(* IEC 61131-3 sources: 89152_FlorisHendrix_AfstudeerProject/89152_FlorisHendrix_ExamenProject/Stations/MachineControl/MachineControl/Class/HwControl, 1 file *)

(* ---- HwControl.st ---- *)
#include "..\..\Class\HwControl\HwControl.h"
#include "..\..\Class\HwControl\watchdog.h"
#include "..\..\Source\interfaces\lsl_st_sysinfo.h"
#include "..\..\Source\interfaces\lsl_st_systrace.h"
#include "..\..\Class\HwControl\_HWKScope.h"

(*!
<Class
	Name               = "HwControl"
	Revision           = "5.21"
	RealtimeTask       = "false"
	DefRealtime        = "1 ms"
	DefRealtimeIndex   = "0"
	CyclicTask         = "false"
	DefCyclictime      = "1 ms"
	DefCyclicIndex     = "2147483392"
	BackgroundTask     = "false"
	Sigmatek           = "true"
	OSInterface        = "false"
	HighPriority       = "false"
	Automatic          = "false"
	UpdateMode         = "Prescan"
	IconPath           = ".\Class\HwControl\HwControl.ico"
	SharedCommandTable = "true"
	Objectsize         = "(646,120)"
	Comment            = "Class to handle VaranManager,  and the cooperation with DiasMasterC">
	<Channels>
		<Server Name="Control">
		</Server>
		<Server Name="DiasMaster" WriteProtected="false" Comment="connect to client &apos;to_HWControl&quot; of class DiasMasterC if used (if Server is 1 class is connected)&#13;&#10;">
		</Server>
		<Server Name="SafetyState" Visualized="true" Initialize="false" WriteProtected="true" Retentive="false" Comment="Shows state of safety functionality initialisation&#13;&#10;&#13;&#10; 1..OK&#13;&#10; 0..not active or initializing&#13;&#10;-1..failed to allocate memory&#13;&#10;-2..invalid domain number set in this system&#13;&#10;-3..newer OS version required for domain number support&#13;&#10;-4..method to determine domain number not provided by lsl_st_hardwaretree.h&#13;&#10;-5..only 1 instance of safety manager allowed&#13;&#10;-6..a slave system can only have 1 master. check hw class configuration&#13;&#10;-7..invalid module type tried to log in&#13;&#10;-8..couldn&apos;t find InterfaceCRC which is requested by other domain. Check SafetyDesigner projects, most likely the interface variables doesn&apos;t match.&#13;&#10;-9..failed to add a new copy data object to varan manager&#13;&#10;-10..a non-optional module or domain is not available&#13;&#10;-11..timeout in initialisation (see debugger trace or logfile for further details)&#13;&#10;-13..the class safetymanager could not login into the class HwControl."/>
		<Client Name="HwcLogging" Required="true" Internal="true"/>
		<Client Name="HWRtPostScan" Required="true" Internal="true"/>
		<Client Name="InterfaceNo" Required="false" Internal="false" DefValue="1" Comment="If interface frames via IP address are used, this is the place to choose the interface number&#13;&#10;&#13;&#10;For example if you set the IP of interface 1 via autoexec.lsl setting SET IP 1 HOSTADDR x.x.x.x and this is what you want to use, you choose 1 for the interface number."/>
		<Client Name="RtTaskSync" Required="false" Internal="false" DefValue="0" Comment="With this setting the realtime task synchronization between more cores can be activated.&#13;&#10;If it is activated and not supported, the client is set to 0.&#13;&#10;As an initialization value. For further information look at library help.&#13;&#10;0 .. deactivated (default)&#13;&#10;1 .. activated&#13;&#10;&#13;&#10;"/>
		<Client Name="SafetyDomainTimeout" Required="false" Internal="false" Comment="[ms] the class has to wait for optional interface domains (leave 0 if none available)&#13;&#10;Set this client to 1 when using FlexCon functionality (without interface domains) where it&apos;s possible that not all participants are available at all times"/>
		<Client Name="SafetyManager" Required="true" Internal="true"/>
		<Client Name="UdpSafetyPort" Required="false" Internal="false" DefValue="10823" Comment="If interface frames via IP address are used, this is the place to choose the port.&#13;&#10;It&apos;s recommended to only change the port (all communication partners must use the same port!) if there would be a conflict with the default port 10823."/>
	</Channels>
	<Dependencies>
		<Files>
			<File Path=".\Class\VaranManager_Base\VaranManager_Base.h" Include="false"/>
			<File Path=".\Class\HwControl\HwControl.h" Include="true"/>
			<File Path=".\Class\HwControl\watchdog.h" Include="true"/>
			<File Path=".\Source\interfaces\lsl_st_sysinfo.h" Include="true"/>
			<File Path=".\Source\interfaces\lsl_st_systrace.h" Include="true"/>
			<File Path=".\Class\HwControl\_HWKScope.h" Include="true"/>
		</Files>
	</Dependencies>
	<RevDoku>
		<Owner Company="Sigmatek" Author="renste"/>
		<Dokumentation Revision="5.21" Date="30.09.2022" Author="RamAnd" Company="Sigmatek" Description="The busy state of the safety CPU wasn&apos;t detected correctly when establishing UDP connections."/>
		<Dokumentation Revision="5.20" Date="13.07.2022" Author="RamAnd" Company="Sigmatek" Description="Try again to establish a safety UDP connection if the attempt failed because the safe CPU was busy."/>
		<Dokumentation Revision="5.19" Date="22.03.2022" Author="RamAnd" Company="Sigmatek" Description="Added support for the new OS Interface to quit errors"/>
		<Dokumentation Revision="5.18" Date="17.01.2022" Author="EisMic" Company="Sigmatek" Description="Testversion: Forward the NewInst commando CMD_HWC_CONVERT_COMPRESSED_HWPATH to the SafetyManager class."/>
		<Dokumentation Revision="5.17" Date="30.11.2021" Author="EisMic" Company="Sigmatek" Description="Added global functions to determine the current operation system.&#13;&#10;Added global function HWC_IsPostInitFinished to determine if the postinit phase is finished or not."/>
		<Dokumentation Revision="5.16" Date="23.10.2020" Author="PieSte" Company="Sigmatek" Description="Added support for new blocktype and extended routing of FSoE data for this type.&#13;&#10;Corrected allocate of udp buffers at &quot;AddModule()&quot;.&#13;&#10;Don&apos;t Log AddDynSlave error if RetCode is zero at GetDestSafetyOfDO() Methode."/>
		<Dokumentation Revision="5.15" Date="18.12.2020" Author="RamAnd" Company="Sigmatek" Description="Removed CLI/STI occurances in internal time measurements"/>
		<Dokumentation Revision="5.14" Date="13.03.2020" Author="Berste1" Company="Sigmatek" Description="Registration for Pll readjustment added"/>
		<Dokumentation Revision="5.13" Date="08.04.2020" Author="PieSte" Company="Sigmatek" Description="Add client RtTaskSync for realtime synchronization if more than one core is used.&#13;&#10;Corrected nil pointer &quot;pStr_HWTreeEntry&quot; at newinst command &quot;CMD_GET_HARDWARE_DIAGNOSIS&quot;."/>
		<Dokumentation Revision="5.12" Date="02.03.2020" Author="FurDom" Company="Sigmatek" Description="Reworked to support newer CPUs (address space &gt; 0x80000000). Needs SafetyUDP class version &gt;= 1.4!"/>
		<Dokumentation Revision="5.11" Date="14.08.2019" Author="LanSte" Company="Sigmatek" Description="Added header file: _HWKScope.h for scope interface. "/>
		<Dokumentation Revision="5.10" Date="08.11.2019" Author="RamAnd" Company="Sigmatek" Description="Detached the logging functionality from HwControl into a new class HwcLogging which is used now as an embedded object in HwControl.&#13;&#10;Added more logging possibilities via new function _HwcLog_sprintfST."/>
		<Dokumentation Revision="5.9" Date="18.07.2019" Author="RamAnd" Company="Sigmatek" Description="Corrected that SDO forwarding would not work properly in some cases.&#13;&#10;Prevent writing to an invalid pointer when resetting UDP connections that could have lead to a crash."/>
		<Dokumentation Revision="5.8" Date="25.06.2019" Author="RamAnd" Company="Sigmatek" Description="Added support for FlexCon functionality."/>
		<Dokumentation Revision="5.7" Date="14.03.2019" Author="RamAnd" Company="Sigmatek" Description="Removed limitations of formerly unallowed safety topologies (since v4.0)"/>
		<Dokumentation Revision="5.6" Date="12.02.2019" Author="PieSte" Company="Sigmatek" Description="The Sequence Number in the SafetyManager class for Udp Safety communication has been extended from 1 to 4 bytes. This increases the availability of the Udp Safety connection. Furthermore two clients have been added at internal class SafetyManager to set the Request Cycle (Default 10) and the Response Timeout (Default 100ms) to optimize the Safety UDP bus load. This setting may only be changed after consultation with Sigmatek.  (SA43141)&quot;/&gt;"/>
		<Dokumentation Revision="5.5" Date="22.01.2019" Author="EisMic" Company="Sigmatek" Description="Corrected an error that the Realtime/Cyclic task of the class was called 2 times if the derivation of the class has a configured Realtime/Cyclic Task. (The error apperared since v5.0)"/>
		<Dokumentation Revision="5.4" Date="15.11.2018" Author="LanSte" Company="Sigmatek" Description="SafetyManager: Added support for custom FSoE Connections."/>
		<Dokumentation Revision="5.3" Date="27.08.2018" Author="PieSte" Company="Sigmatek" Description="Behaviour of safety udp communication when resetting the bSequenceCntReceived flag after maximum of retries corrected. (SafetyManager)"/>
		<Dokumentation Revision="5.2" Date="18.07.2018" Author="PieSte&#13;&#10;EisMic" Company="Sigmatek" Description="Added support for HGW1033-3. (in SafetyManager)&#13;&#10;Removed incorrect LogMessage. Corrected access exception in method CalculateTaskInfo.&#13;&#10;OS_AddTraceKeyVal is not used anymore with OS-Version between 9.1.0 and 9.3.0. Not supported with these versions."/>
		<Dokumentation Revision="5.1" Date="19.06.2018" Author="ZoePat" Company="Sigmatek" Description="Corrected a possible reboot of some CPUs (CCP512, CCP612, CP212, and similar). The error appeared since V5.0 if the SRAM was accessed via the cyclic-task of the HWControl."/>
		<Dokumentation Revision="5.0" Date="26.03.2018" Author="EisMic" Company="Sigmatek" Description="Added support for 2nd realtime.&#13;&#10;Added support for 2nd varanmanager.&#13;&#10;Removed task settings from object. Task-settings for realtime and cyclic task are now calculated depending on the connected hardware-classes. See documentation for more details.&#13;&#10;Extended the methods AddFirstCallHw and AddHwObject by some parameters to select a CPU-core and task-times.&#13;&#10;Added support for SmartIO modules."/>
		<Dokumentation Revision="4.15" Date="06.03.2018" Author="EisMic" Company="Sigmatek" Description="Attached header files no longer point to the installation directory of LASAL but instead now point to the the source/interfaces folder."/>
		<Dokumentation Revision="4.14" Date="18.01.2018" Author="EisMic" Company="Sigmatek" Description="Added new NewInst command to get supported features by HwControl.&#13;&#10;The newinst cmd CMD_SET_POSTINIT_DONE will now be send to all connected classes instead of only to the DiasMaster."/>
		<Dokumentation Revision="4.13" Date="23.01.2018" Author="RamAnd" Company="Sigmatek" Description="Log messages have been standardized for easier maintenance, easier use in any class and to allow spam filtering. Code for the logging functions is now only located in HwControl."/>
		<Dokumentation Revision="4.12" Date="05.01.2018" Author="PieSte" Company="Sigmatek" Description="The safety UDP communication at &quot;SafetyManager&quot; class has been made more reliable. Now only new packages are allowed and old packages are discarded."/>
		<Dokumentation Revision="4.11" Date="18.09.2017" Author="LanSte" Company="Sigmatek" Description="Added NewInst Commands to check if the Post-Init is done."/>
		<Dokumentation Revision="4.10" Date="29.08.2017" Author="RamAnd" Company="Sigmatek" Description="The VaranManager can now tell the HwControl if it doesn&apos;t have any clients connected. In this case the HwControl is in charge of triggering the internal watchdog."/>
		<Dokumentation Revision="4.9" Date="22.08.2017" Author="RamAnd" Company="Sigmatek" Description="Fixed an error which prevented two SCP111s on the same PLC from exchanging interfaceframes in both directions."/>
		<Dokumentation Revision="4.8" Date="23.05.2017" Author="RamAnd" Company="Sigmatek" Description="A pointer for dynamic parameters has been added to the hardware diagnosis. Added initialisation of the pointer with NIL."/>
		<Dokumentation Revision="4.7" Date="22.06.2017" Author="RamAnd" Company="Sigmatek" Description="If a disconnect happens in a multi master system with safety communication (more than 2 systems connected and exchanging safety data) now the other masters are notified about it to reestablish the connection."/>
		<Dokumentation Revision="4.6" Date="01.03.2017" Author="EisMic" Company="Sigmatek" Description="Corrected an error in the handling of optional safety modules."/>
		<Dokumentation Revision="4.5" Date="14.02.2017" Author="ZoePat" Company="Sigmatek" Description="SdiasModules can now request to increase the PostInit timeout."/>
		<Dokumentation Revision="4.4" Date="21.09.2016" Author="PieSte" Company="Sigmatek" Description="Add methode &quot;AddFirstCallHW&quot; for objects which are called as first at HwControl Realtime. In the TraceView scope is the and of first object call as UserEvent0 with data = 1.215.775.599 marked. "/>
		<Dokumentation Revision="4.3" Date="28.01.2016" Author="RamAnd" Company="Sigmatek" Description="Support for FSoE via IP added."/>
		<Dokumentation Revision="4.2" Date="06.06.2016" Author="EisMic" Company="Sigmatek" Description="Corrected error if distributed safety modules are connected after the initialisation phase."/>
		<Dokumentation Revision="4.1" Date="11.05.2016" Author="RamAnd" Company="Sigmatek" Description="Suppressed warning that would occur with target ARM on compiler version 30 or higher."/>
		<Dokumentation Revision="4.0" Date="30.11.2015" Author="ZoePat&#13;&#10;LanSte" Company="Sigmatek" Description="Check for unallowed safety topology."/>
		<Dokumentation Revision="3.9" Date="21.10.2015" Author="RamAnd" Company="Sigmatek" Description="Support for MS012 added"/>
		<Dokumentation Revision="3.8" Date="19.05.2015" Author="RamAnd" Company="Sigmatek" Description="If two systems with FSoE safety were connected via VBC/VMC an error in the connection establishment could cause the FSoE connection to fail."/>
		<Dokumentation Revision="3.7" Date="15.04.2015" Author="RamAnd" Company="Sigmatek" Description="Added another step in initialisation to prevent watchdog error."/>
		<Dokumentation Revision="3.6" Date="16.10.2014&#13;&#10;25.03.2015" Author="RamAnd&#13;&#10;PieSte" Company="Sigmatek" Description="Support for SCP111 added.&#13;&#10;Support for SDD1300, SDD1400, SDD1500 and SDD1600 added."/>
		<Dokumentation Revision="3.5" Date="12.11.2014" Author="PieSte" Company="Sigmatek" Description="Removed trace message if watchdog interface is not available."/>
		<Dokumentation Revision="3.4" Date="28.10.2014" Author="RamAnd" Company="Sigmatek" Description="If an error has been reported to HwControl, it is now forwarded to the DiasMasterC object (if there is one)."/>
		<Dokumentation Revision="3.3" Date="10.10.2014" Author="PieSte" Company="Sigmatek" Description="Added Watchdog API and trigger watchdog in postscan task."/>
		<Dokumentation Revision="3.2" Date="18.06.2014" Author="EisMic" Company="Sigmatek" Description="Added support for reading hardware diagnosis via newinst cmd: CMD_GET_HARDWARE_DIAGNOSE "/>
		<Dokumentation Revision="3.1" Date="17.06.2014" Author="RamAnd" Company="Sigmatek" Description="Added possibility to start a quit error via OS interface."/>
		<Dokumentation Revision="3.0" Date="15.04.2014" Author="RamAnd" Company="Sigmatek" Description="Changed initialisation: &#13;&#10; - Activation of hardware classes realtime task as well as completing CDIAS/DIAS initialisation is now done in post init instead of last init&#13;&#10; - No realtime is running in the first initialisation of the modules&#13;&#10; - New second initialisation where realtime is running to check if the realtime data are valid"/>
		<Dokumentation Revision="2.0" Date="12.02.2014" Author="PieSte" Company="Sigmatek" Description="Improved description of CyWork method."/>
		<Dokumentation Revision="1.50" Date="06.12.2013" Author="LanSte&#13;&#10;RamAnd&#13;&#10;FucHer" Company="Sigmatek" Description="Ensured that he class is copatible with old loader versions that do not support the post init phase.&#13;&#10;Removed domain support&#13;&#10;Changed AWL code to Structured Text.&#13;&#10;If the task setting for cyclic task fails, the error wasn&apos;t displayed.&#13;&#10;The task setting for cyclic task didn&apos;t work (only required if existing object is updated)."/>
		<Dokumentation Revision="1.40" Date="01.08.2013" Author="RamAnd" Company="Sigmatek" Description="Corrected error, where the user classes are already called during SDIAS initialisation."/>
		<Dokumentation Revision="1.30" Date="18.07.2013" Author="RamAnd" Company="Sigmatek" Description="Added PostInit interface of loader, where after the last init the varan managers can initialize modules until they are ready."/>
		<Dokumentation Revision="1.20" Date="07.03.2013" Author="RamAnd" Company="Sigmatek" Description="Changed range of the safety NewInst commands. Range for HW-Classes: 0x8000-0x8FFF; Range for Safety HW-Classes: 0x8100-0x81FF"/>
		<Dokumentation Revision="1.15" Date="23.12.2011" Author="RamAnd" Company="Sigmatek" Description="Added support for the SafetyManager"/>
		<Dokumentation Revision="1.14" Date="14.02.2012" Author="RamAnd" Company="Sigmatek" Description="Watchdog is now also triggered if no VARAN/DIAS interface is available (needed for internal IOs of Edge ETVs)"/>
		<Dokumentation Revision="1.13" Date="25.05.2011" Author="RamAnd" Company="Sigmatek" Description="PostScan-Calls in Init-Phase are now done in HwControl instead of VaranManager."/>
		<Dokumentation Revision="1.12" Date="27.10.2010" Author="RamAnd" Company="Sigmatek" Description="Added RtPostScan support for special hardware like the IOs of an Edge ETV"/>
		<Dokumentation Revision="1.11" Date="13.08.2010" Author="BleErn" Company="Sigmatek" Description="Postscan calls were not stopped on error"/>
		<Dokumentation Revision="1.10" Date="22.07.2010" Author="WocPet" Company="Sigmatek" Description="New functionality added to display required error from diasmaster"/>
		<Dokumentation Revision="1.9" Date="13.07.2010" Author="BleErn" Company="Sigmatek" Description="Content of corresponding LASAL Hardware Description file (.lhd) which is necessary for the hardware editor has been corrected"/>
		<Dokumentation Revision="1.8" Date="03.03.2010" Author="BleErn" Company="Sigmatek" Description="Added Handling for DiasMaster RtPostScan"/>
		<Dokumentation Revision="1.7" Date="08.02.2010" Author="BleErn" Company="Sigmatek" Description="Added Baseclass for RtPostScan with DIAS/CDIAS/CTMS&#13;&#10;Caution: RtPostScan cannot be used together with RtDebug!"/>
		<Dokumentation Revision="1.6" Date="10.03.2010" Author="RamAnd" Company="Sigmatek" Description="Added Support for various IOs (e.g. ETV Edge IOs)"/>
		<Dokumentation Revision="1.5" Date="03.02.2009" Author="RamAnd" Company="Sigmatek" Description="Added Synchronity check if VMC is used."/>
	</RevDoku>
	<Network Name="HwControl">
		<!-- List of Components in this network -->
		<Components>
			<Object
				Name       = "_base"
				Class      = "HwControlBase"
				Position   = "(218,120)"
				Visualized = "false"
				RealTime   = "1 ms">
				<Channels>
					<Server Name="Control"/>
					<Server Name="DiasMaster"/>
					<Server Name="State"/>
					<Client Name="RtDebug"/>
					<Client Name="To_StdLib"/>
					<Client Name="To_TaskObjectControl"/>
				</Channels>
			</Object>
			<Object
				Name       = "HwcLogging"
				Class      = "HwcLogging"
				Position   = "(150,540)"
				Visualized = "false">
				<Channels>
					<Server Name="ClassSvr"/>
					<Server Name="OverrideSpamProtection"/>
					<Client Name="To_SigCLib"/>
				</Channels>
			</Object>
			<Object
				Name       = "HWRtPostScan"
				Class      = "HWRtPostScan"
				Position   = "(150,930)"
				Visualized = "false"
				RealTime   = "1 ms"
				RealIndex  = "1073741824">
				<Channels>
					<Server Name="ClassSvr"/>
					<Client Name="toHwControlBase"/>
				</Channels>
			</Object>
			<Object
				Name       = "SafetyManager"
				Class      = "SafetyManager"
				Position   = "(960,360)"
				Visualized = "true"
				CyclicTime = "10 ms">
				<Channels>
					<Server Name="ClassState"/>
					<Server Name="InitFault"/>
					<Server Name="InitSSM"/>
					<Server Name="LoginCnt"/>
					<Server Name="MaxSyncDuration"/>
					<Server Name="MinSyncDuration"/>
					<Server Name="sControl"/>
					<Server Name="sErrorCount"/>
					<Server Name="sLastErrorMessage"/>
					<Server Name="sLastErrorNoOS"/>
					<Server Name="sTReceive"/>
					<Server Name="SyncDuration"/>
					<Client Name="InterfaceNo" Value="1"/>
					<Client Name="SafetyDomainTimeout"/>
					<Client Name="To_HwControl"/>
					<Client Name="To_MultiTask"/>
					<Client Name="To_OSKernel"/>
					<Client Name="UdpSafetyPort" Value="10823"/>
					<Client Name="UdpSafetyRequestCycle" Value="UDP_MIN_REQUEST_TIME"/>
					<Client Name="UdpSafetyResponseTimeout" Value="UDP_MIN_RESPONSE_TIMEOUT"/>
				</Channels>
			</Object>
		</Components>
		<Comments>
		</Comments>
		<!-- List of Connections in this network -->
		<Connections>
			<Connection Source="this.Control" Destination="_base.Control" Vertices="(1794,210),(886,210),"/>
			<Connection Source="this.State" Destination="_base.State" Vertices="(1794,270),(886,270),"/>
			<Connection Source="this.DiasMaster" Destination="_base.DiasMaster" Vertices="(1794,330),(886,330),"/>
			<Connection Source="_base.RtDebug" Destination="this.RtDebug" Vertices="(218,330),(120,330),(120,210),(38,210),"/>
			<Connection Source="this.SafetyManager" Destination="SafetyManager.ClassState"/>
			<Connection Source="SafetyManager.To_HwControl" Destination="_base.Control" Vertices="(960,570),(930,570),(930,210),(886,210),"/>
			<Connection Source="SafetyManager.UdpSafetyPort" Destination="this.UdpSafetyPort" Vertices="(960,450),(38,450),"/>
			<Connection Source="SafetyManager.SafetyDomainTimeout" Destination="this.SafetyDomainTimeout" Vertices="(960,750),(930,750),(930,750),(120,750),(120,390),(38,390),"/>
			<Connection Source="SafetyManager.InterfaceNo" Destination="this.InterfaceNo" Vertices="(960,510),(38,510),"/>
			<Connection Source="this.SafetyState" Destination="SafetyManager.ClassState" Vertices="(1794,390),(1740,390),(1740,450),(1622,450),"/>
			<Connection Source="this.HWRtPostScan" Destination="HWRtPostScan.ClassSvr"/>
			<Connection Source="HWRtPostScan.toHwControlBase" Destination="_base.Control" Vertices="(150,1020),(120,1020),(120,870),(930,870),(930,210),(886,210),"/>
			<Connection Source="this.HwcLogging" Destination="HwcLogging.ClassSvr"/>
		</Connections>
		<!-- Headerfiles -->
		<Options>
		</Options>
	</Network>
</Class>
*)
#pragma using HwControlBase

HwControl : CLASS
: HwControlBase
	TYPE
	  pVaranManager : ^VaranManager;
	  t_DMFunctions : STRUCT
	    p_RtFunction : pVoid;
	    p_SendSync : pVoid;
	    p_FinishIMProg : pVoid;
	    p_LastInit : pVoid;
	    p_This : pVoid;
	    sd_PllTime : DINT;
	    ud_DiasTime : UDINT;
	    sd_RtDebug : DINT;
	    p_RtPostScanFunction : pVoid;
	    SafetyManagerThisPointer : ^pVirtualBase;
	  END_STRUCT;
	  t_DiasMaster : STRUCT
	    ud_Counter : UDINT;
	    p_Functions : ^t_DMFunctions;
	  END_STRUCT;
#pragma pack(push, 1)
	  t_HwObjectListCallFirst : STRUCT
	    pThis : pVirtualBase;
	    udLoggedInNumber : UDINT;
	    us_CoreSelect : USINT;
	    ud_RtTime_us : UDINT;
	    ud_CyTime_us : UDINT;
	    pNext : ^t_HwObjectListCallFirst;
	  END_STRUCT;
#pragma pack(pop)
#pragma pack(push, 1)
	  t_HwObjectListElement : STRUCT
	    pThis : pVirtualBase;
	    pRtPostScan : ^UDINT;  //! <Type Comment="used for EdgeETV IOs" Name="t_HwObjectListElement.pRtPostScan"/>
	    bdSettings : t_HwObjListSettings;
	    usEscSequence : USINT;  //! <Type Comment="Escapesequence that identifies the bustype." Name="t_HwObjectListElement.usEscSequence"/>
	    us_CoreSelect : USINT;
	    ud_RtTime_us : UDINT;
	    ud_CyTime_us : UDINT;
	    pNext : ^t_HwObjectListElement;
	  END_STRUCT;
#pragma pack(pop)
	  t_VMFunctions : STRUCT
	    p_This : pVaranManager;
	    ud_VaranTime : UDINT;
	    b_IsAlsoClient : BOOL;
	    ud_SuperiorTime : UDINT;
	    b_HWClassSynchron : BOOL;
	    b_OverrideFrameCheck : BOOL;
	    SafetyManagerThisPointer : ^pVirtualBase;
	    Reserved1 : DINT;
	    Reserved2 : DINT;
	  END_STRUCT;
	  t_OneVaranManager : STRUCT
	    ud_CounterRt : UDINT;
	    ud_CounterCy : UDINT;
	    ud_SuperiorSync : UDINT;
	    ud_SuperiorSyncActual : UDINT;
	    p_Functions : ^t_VMFunctions;
	    usOldFrameCnt : USINT;
	    usActFrameCnt : USINT;
	    usSyncCheck : USINT;
	    us_CoreSelect : USINT;
	    ud_RtTime_us : UDINT;
	    ud_CyTime_us : UDINT;
	  END_STRUCT;
#pragma pack(push, 1)
	  t_s_CallFirstObject : STRUCT
	    pThis : pVirtualBase;
	    us_CoreSelect : USINT;
	    ud_RtTime_us : UDINT;
	    ud_CyTime_us : UDINT;
	  END_STRUCT;
#pragma pack(pop)
#pragma pack(push, 1)
	  t_s_RtTaskControl : STRUCT
	    pvPreRtSyncTaskEvent : pVoid;
	    pvPostRtSyncTaskEvent : pVoid;
	    udPreRtCnt : UDINT;
	    udPostRtCnt : UDINT;
	    b_RtTaskControlActive : BOOL;
	    usCoresRtActive : USINT;
	  END_STRUCT;
#pragma pack(pop)
#pragma pack(push, 1)
	  t_s_TaskCoreInfo : STRUCT
	    us_CoreSelect : USINT;
	    ud_MyRtTaskTime_us : UDINT;  //! <Type Comment="tasktime of HwControl realtime task of the core" Name="t_s_TaskCoreInfo.ud_MyRtTaskTime_us"/>
	    ud_MyCyTaskTime_us : UDINT;  //! <Type Comment="tasktime of HwControl cyclic task of the core" Name="t_s_TaskCoreInfo.ud_MyCyTaskTime_us"/>
	    uiHwTimeStamp_us : UINT;
	    ud_FirstPostScanCall : UDINT;
	    ud_LastPostScanWorkCall : UDINT;
	    b_PostScanStarted : BOOL;
	  END_STRUCT;
#pragma pack(pop)
	END_TYPE
  //Servers:
	SafetyState 	: SvrCh_DINT;
  //Clients:
	SafetyManager 	: CltChCmd_SafetyManager;
	SafetyDomainTimeout 	: CltCh_UDINT;
	UdpSafetyPort 	: CltCh_UDINT;
	InterfaceNo 	: CltCh_UDINT;
	RtTaskSync 	: CltCh_DINT;
	HWRtPostScan 	: CltChCmd_HWRtPostScan;
	HwcLogging 	: CltChCmd_HwcLogging;
  //Variables:
		a_VaranManager : ARRAY [0..MAX_VARAN_MANAGERS-1] OF t_OneVaranManager;
			//! <Variable Comment="array of structures for VaranManager functions and settings" Name="a_VaranManager"/>
		s_DiasMaster 	: t_DiasMaster;			//! <Variable Comment="structure for DiasMaster functions and settings" Name="s_DiasMaster"/>
		us_Initcounter 	: USINT;			//! <Variable Comment="varaiable to count init steps" Name="us_Initcounter"/>
		p_DebugAPI 	: ^DEBUGAPI;			//! <Variable Comment="pointer to debug API (OS - Interface)" Name="p_DebugAPI"/>
		p_WatchdogAPI 	: ^LSLAPI_IWATCHDOG;
		pCallFirstObjects 	: ^t_HwObjectListCallFirst;
		sCallFirstObjects : ARRAY [0..HWCONTROL_MAX_FIRSTCALL_OBJECTS-1] OF t_s_CallFirstObject;

		bCallFirstObjects 	: BOOL;
		VaranManagersAvailable 	: USINT;
		pSCDW 	: ^LSL_CDIASWATCHDOG;
		pHwControlLogins 	: ^t_HwObjectListElement;
		b_PostInitInstalled 	: BOOL;
		pSystrace 	: ^OS_SYSTRACE;
		AdditionalPostInitTime 	: UDINT;
		SupportedFeatures 	: t_HWC_SupportedFeatureBits1;
		pLSLSysInfo 	: ^LSL_SYSINFO_TYPE;
		ud_CPUCoreCount 	: UDINT;			//! <Variable Comment="Shows the amount of CPU cores of the current CPU." Name="ud_CPUCoreCount"/>
		us_CPUsRtCyEnabled 	: USINT;
		aHwControl_Times : ARRAY [0..TASK_SELECT_COREMAX] OF t_HwControl_Times_SINGLE;
			//! <Variable Comment="Shows the measured times if the time measurement is activated in HwControl.h with the define HWCONTROL_TIME_MEASUREMENT." Name="aHwControl_Times"/>
		aTaskInfoCore : ARRAY [0..TASK_SELECT_COREMAX] OF t_s_TaskCoreInfo;
			//! <Variable Comment="Shows information of the supported cores." Name="aTaskInfoCore"/>
		sRtTaskControl 	: t_s_RtTaskControl;
		pSpecialObjects 	: ^t_HwObjectListElement;
		mt_api 	: ^LSL_MT_TYPE;
		b_SoftwareSyncActive 	: BOOL;
  //Functions:
				//! <Function Comment="[#ENGLISH]&#13;&#10;=================================================================================================&#13;&#10;Init for HwControl class&#13;&#10;=================================================================================================&#13;&#10;[clients] RtDebug    :R&#13;&#10;[members] us_InitCounter  :R/W :varaiable to count init steps&#13;&#10;   p_DebugAPI   :W  :pointer to debug API (OS - Interface)&#13;&#10;   s_DiasMaster  :R  :structure for DiasMaster functions and settings&#13;&#10;" Name="Init"/>
	FUNCTION VIRTUAL GLOBAL Init;

	FUNCTION VIRTUAL GLOBAL CyWork
		VAR_INPUT
			EAX 	: UDINT;
		END_VAR
		VAR_OUTPUT
			state (EAX) 	: UDINT;
		END_VAR;

	FUNCTION VIRTUAL GLOBAL RtWork
		VAR_INPUT
			EAX 	: UDINT;
		END_VAR
		VAR_OUTPUT
			state (EAX) 	: UDINT;
		END_VAR;

	FUNCTION HwControl
		VAR_OUTPUT
			ret_code 	: ConfStates;
		END_VAR;

	FUNCTION VIRTUAL GLOBAL UpdateRtPostScan;
				//! <Function Comment="no longer used." Name="AddSafetyManager"/>
	FUNCTION VIRTUAL GLOBAL AddSafetyManager
		VAR_INPUT
			pThis 	: pVirtualBase;
		END_VAR
		VAR_OUTPUT
			pFirstVM 	: pVirtualBase;
		END_VAR;
				//! <Function Comment="no longer used." Name="DisableSafetyManager"/>
	FUNCTION VIRTUAL GLOBAL DisableSafetyManager;
				//! <Function Comment="[#ENGLISH]&#13;&#10;=================================================================================================&#13;&#10;Class to call a function pointer&#13;&#10;=================================================================================================&#13;&#10;" Name="CallPtr"/>
	FUNCTION CallPtr
		VAR_INPUT
			p_function 	: pVoid;			//! <Variable Comment="pointer to function should be called" Name="CallPtr.p_function"/>
			p_this 	: pVoid;			//! <Variable Comment="thispointer of object" Name="CallPtr.p_this"/>
		END_VAR;
				//! <Function Comment="Function to get Tasktime of Hwcontrol class&#13;&#10;" Name="GetMyTaskTime"/>
	FUNCTION GLOBAL GetMyTaskTime
		VAR_INPUT
			us_CoreSelect 	: DINT := 0;			//! <Variable Comment="Coreselect 0 ... ud_task_time is realtime task time of core 0.&#13;&#10;Coreselect 1 ... ud_task_time is realtime task time of core 1." Name="GetMyTaskTime.us_CoreSelect"/>
		END_VAR
		VAR_OUTPUT
			ud_task_time 	: UDINT;			//! <Variable Comment="rt task time in ns" Name="GetMyTaskTime.ud_task_time"/>
		END_VAR;
				//! <Function Comment="Function to add a VaranManager to HwControl list" Name="AddVaranManager"/>
	FUNCTION GLOBAL AddVaranManager
		VAR_INPUT
			ud_manager_number 	: UDINT;			//! <Variable Comment="number of varan manager&#13;&#10;" Name="AddVaranManager.ud_manager_number"/>
			p_function_list 	: ^void;			//! <Variable Comment="pointer to function list and settings of VaranMaster" Name="AddVaranManager.p_function_list"/>
			us_CoreSelect 	: USINT := 0;			//! <Variable Comment="Selection on which core the manager should be called." Name="AddVaranManager.us_CoreSelect"/>
			ud_RtTime_us 	: UDINT := 0;			//! <Variable Comment="Realtime task time in µs.&#13;&#10;The time will be used in the calculation for the realtime task time of the selected core.&#13;&#10;The calculated time of the HwControl will be distributed to the logged in object with the newinst command CMD_POST_INIT_DISTRIBUTE_TASKTIMES.&#13;&#10;For more information about the task time settings look in the hardware class documentation." Name="AddVaranManager.ud_RtTime_us"/>
			ud_CyTime_us 	: UDINT := 0;			//! <Variable Comment="Cyclic task time in µs.&#13;&#10;The time will be used in the calculation for the cyclic task time of the selected core.&#13;&#10;The calculated time of the HwControl will be distributed to the logged in object with the newinst command CMD_POST_INIT_DISTRIBUTE_TASKTIMES.&#13;&#10;For more information about the task time settings look in the hardware class documentation." Name="AddVaranManager.ud_CyTime_us"/>
		END_VAR
		VAR_OUTPUT
			sd_retval 	: DINT;			//! <Variable Comment="Returncode of the function.&#13;&#10;0 ... OK&#13;&#10;&lt;&gt; 0 ... Error" Name="AddVaranManager.sd_retval"/>
		END_VAR;
				//! <Function Comment="Function to remove a Varanmanager from the HwControl list." Name="DisableVaranManager"/>
	FUNCTION GLOBAL DisableVaranManager
		VAR_INPUT
			ud_manager_number 	: UDINT;			//! <Variable Comment="number of varan manager" Name="DisableVaranManager.ud_manager_number"/>
			p_function_list 	: ^void;			//! <Variable Comment="pointer to function list and settings of VaranMaster" Name="DisableVaranManager.p_function_list"/>
		END_VAR
		VAR_OUTPUT
			sd_retval 	: DINT;			//! <Variable Comment="Returncode of the function.&#13;&#10;0 ... OK&#13;&#10;&lt;&gt; 0 ... Error" Name="DisableVaranManager.sd_retval"/>
		END_VAR;
				//! <Function Comment="Function sets Hardware off&#13;&#10;" Name="SetHardwareOff"/>
	FUNCTION GLOBAL SetHardwareOff
		VAR_INPUT
			e_error 	: t_e_VaranErrors;			//! <Variable Comment="reason why hardware is set off" Name="SetHardwareOff.e_error"/>
		END_VAR;
				//! <Function Comment="Function returns Debug State" Name="GetRtDebugState"/>
	FUNCTION GLOBAL GetRtDebugState
		VAR_OUTPUT
			sd_RtDebug 	: DINT;
		END_VAR;
				//! <Function Comment="function to add a special hw. &#13;&#10;function should only be used from hardware classes.&#13;&#10;Has to be called in initialisation phase.&#13;&#10;&#13;&#10;This object will be called in realtime and cyclic task from the HwControl. Only on core 0.&#13;&#10;&#13;&#10;Attention:&#13;&#10;To select a core on which the special hw should be called, please use the method AddHwObject." Name="AddSpecialHW"/>
	FUNCTION GLOBAL AddSpecialHW
		VAR_INPUT
			pThis 	: pVirtualBase;			//! <Variable Comment="Thispointer of object." Name="AddSpecialHW.pThis"/>
			pRtPostScan 	: ^UDINT;
		END_VAR
		VAR_OUTPUT
			retcode 	: DINT;
		END_VAR;

	FUNCTION PostScanWork
		VAR_INPUT
			us_CoreSelect 	: USINT;
		END_VAR;
				//! <Function Comment="This function prototype is used to call functions via function pointers." Name="ObjectFunct"/>
	FUNCTION ObjectFunct;
				//! <Function Comment="function to login objects which are called as first objects in HwControl realtime.&#13;&#10;Has to be called in initialisation phase.&#13;&#10;&#13;&#10;Objects which are logged in at the HwControl via this function will get an NewInst call with the command CMD_POST_INIT_DISTRIBUTE_TASKTIMES at the beginning of the post init phase.&#13;&#10;The calculated tasktimes (realtime and cyclic) will be distributed to the classes. The data structure of the command can be seen at the definition of the NewInst command in the Headerfile HwControl.h." Name="AddFirstCallHW"/>
	FUNCTION GLOBAL AddFirstCallHW
		VAR_INPUT
			pThis 	: pVirtualBase;			//! <Variable Comment="pointer on object to call in RtWork" Name="AddFirstCallHW.pThis"/>
			udSelectPlace 	: UDINT;			//! <Variable Comment="Select order of first calls beginning from 0.&#13;&#10;Only one number per object possible.&#13;&#10;0 .. first object&#13;&#10;1 .. second object&#13;&#10;2 .. third object&#13;&#10;....&#13;&#10;max place .. last object" Name="AddFirstCallHW.udSelectPlace"/>
			us_CoreSelect 	: USINT := 0;			//! <Variable Comment="Selection from which core the object should be called.&#13;&#10;0 ... Core 0&#13;&#10;1 ... Core 1&#13;&#10;x ... Core x" Name="AddFirstCallHW.us_CoreSelect"/>
			ud_RtTime_us 	: UDINT := 0;			//! <Variable Comment="Realtime task time in µs.&#13;&#10;The time will be used in the calculation for the realtime task time of the selected core.&#13;&#10;The calculated time of the HwControl will be distributed to the logged in object with the newinst command CMD_POST_INIT_DISTRIBUTE_TASKTIMES.&#13;&#10;For more information about the task time settings look in the hardware class documentation." Name="AddFirstCallHW.ud_RtTime_us"/>
			ud_CyTime_us 	: UDINT := 0;			//! <Variable Comment="Cyclic task time in µs.&#13;&#10;The time will be used in the calculation for the cyclic task time of the selected core.&#13;&#10;The calculated time of the HwControl will be distributed to the logged in object with the newinst command CMD_POST_INIT_DISTRIBUTE_TASKTIMES.&#13;&#10;For more information about the task time settings look in the hardware class documentation." Name="AddFirstCallHW.ud_CyTime_us"/>
		END_VAR
		VAR_OUTPUT
			retcode 	: DINT;			//! <Variable Comment="return value of function&#13;&#10; 0 .. ok&#13;&#10;-1  ... invalid place number&#13;&#10;-2  ... place already selected&#13;&#10;-3  ... object login is to late, it must be done before last init cycle&#13;&#10;-4  ... parameter us_CoreSelect is invalid. (see debugger trace for details)&#13;&#10;-5  ... multicore support not supported by LSL_ITASK interface.&#13;&#10;-6  ... HwControl does not support the number of parameter us_CoreSelect&#13;&#10;-7  ... parameter ud_RtTime_us is smaller than CPU maintimer.&#13;&#10;-8  ... parameter ud_RtTime_us is not a multiple of CPU maintimer.&#13;&#10;-9  ... parameter ud_CyTime_us is smaller than CPU maintimer.&#13;&#10;-10 ... parameter ud_RtTime_us is not a multiple of CPU maintimer." Name="AddFirstCallHW.retcode"/>
		END_VAR;

	FUNCTION InstallPostInitCB
		VAR_OUTPUT
			sd_retval 	: DINT;
		END_VAR;

	FUNCTION UpdateRtFirstCallObjects
		VAR_INPUT
			usCoreSelect 	: USINT;
		END_VAR;

	FUNCTION UpdateRtLoginObjects
		VAR_INPUT
			usCoreSelect 	: USINT;
		END_VAR;

	FUNCTION UpdateRtPostscanLoginObjects
		VAR_INPUT
			usCoreSelect 	: USINT;
		END_VAR;

	FUNCTION UpdateRtVaranManager
		VAR_INPUT
			usActiveCore 	: USINT;
		END_VAR;

	FUNCTION UpdateRtPostScanVaranManager
		VAR_INPUT
			usActiveCore 	: USINT;
		END_VAR;
				//! <Function Comment="function to add a hw object which will be called in the realtime and cyclic task on the selected core.&#13;&#10;function should only be used from hardware classes.&#13;&#10;Has to be called in initialisation phase." Name="AddHwObject"/>
	FUNCTION GLOBAL AddHwObject
		VAR_INPUT
			pThis 	: pVirtualBase;			//! <Variable Comment="Thispointer of object." Name="AddHwObject.pThis"/>
			Settings 	: t_HwObjListSettings;
			EscapeSequence 	: USINT := 0;
			us_CoreSelect 	: USINT := 0;			//! <Variable Comment="Selection from which core the object should be called.&#13;&#10;0 ... Core 0&#13;&#10;1 ... Core 1&#13;&#10;x ... Core x" Name="AddHwObject.us_CoreSelect"/>
			ud_RtTime_us 	: UDINT := 0;			//! <Variable Comment="Realtime task time in µs.&#13;&#10;The time will be used in the calculation for the realtime task time of the selected core.&#13;&#10;The calculated time of the HwControl will be distributed to the logged in object with the newinst command CMD_POST_INIT_DISTRIBUTE_TASKTIMES.&#13;&#10;For more information about the task time settings look in the hardware class documentation." Name="AddHwObject.ud_RtTime_us"/>
			ud_CyTime_us 	: UDINT := 0;			//! <Variable Comment="Cyclic task time in µs.&#13;&#10;The time will be used in the calculation for the cyclic task time of the selected core.&#13;&#10;The calculated time of the HwControl will be distributed to the logged in object with the newinst command CMD_POST_INIT_DISTRIBUTE_TASKTIMES.&#13;&#10;For more information about the task time settings look in the hardware class documentation." Name="AddHwObject.ud_CyTime_us"/>
		END_VAR
		VAR_OUTPUT
			retcode 	: DINT;			//! <Variable Comment="return value of function&#13;&#10; 0 .. ok&#13;&#10;-1  ... failed to allocate memory for hw object&#13;&#10;-2  ... parameter pThis is invalid&#13;&#10;-4  ... parameter us_CoreSelect is invalid. (see debugger trace for details)&#13;&#10;-5  ... multicore support not supported by LSL_ITASK interface.&#13;&#10;-6  ... HwControl does not support the number of parameter us_CoreSelect&#13;&#10;-7  ... parameter ud_RtTime_us is smaller than CPU maintimer.&#13;&#10;-8  ... parameter ud_RtTime_us is not a multiple of CPU maintimer.&#13;&#10;-9  ... parameter ud_CyTime_us is smaller than CPU maintimer.&#13;&#10;-10 ... parameter ud_RtTime_us is not a multiple of CPU maintimer." Name="AddHwObject.retcode"/>
		END_VAR;

	FUNCTION CalcTimeMeasurementPreScan
		VAR_INPUT
			pHwControlTimes 	: ^t_HwControl_Times_SINGLE;
		END_VAR;

	FUNCTION CalcTimeMeasurementPostScan
		VAR_INPUT
			pHwControlTimes 	: ^t_HwControl_Times_SINGLE;
		END_VAR;

	FUNCTION CalcTimeMeasurementCyclic
		VAR_INPUT
			pHwControlTimes 	: ^t_HwControl_Times_SINGLE;
		END_VAR;

	FUNCTION CalculateTaskInfo
		VAR_INPUT
			us_CoreSelect 	: USINT;
			pTaskInfo 	: ^t_s_TaskCoreInfo;
		END_VAR;

	FUNCTION CalculateGGT
		VAR_INPUT
			Var1 	: UDINT;
			Var2 	: UDINT;
		END_VAR
		VAR_OUTPUT
			ggT 	: UDINT;
		END_VAR;

	FUNCTION RtPreScan_CoreX
		VAR_INPUT
			pCoreSelect 	: ^void;
		END_VAR;

	FUNCTION CyWork_CoreX
		VAR_INPUT
			pCoreSelect 	: ^void;
		END_VAR;

	FUNCTION RtPostScan_CoreX
		VAR_INPUT
			pCoreSelect 	: ^void;
		END_VAR;
				//! <Function Comment="Function which returns the ITASK Version of the OS." Name="Get_ITASK_Version"/>
	FUNCTION Get_ITASK_Version
		VAR_OUTPUT
			version 	: UDINT;
		END_VAR;

	FUNCTION VIRTUAL GLOBAL Control::NewInst
		VAR_INPUT
			pPara 	: ^CmdStruct;
			pResult 	: ^results;
		END_VAR
		VAR_OUTPUT
			ret_code 	: iprStates;
		END_VAR;
				//! <Function Comment="[#ENGLISH]&#13;&#10;=================================================================================================&#13;&#10;Write Function of DiasMaster&#13;&#10;=================================================================================================&#13;&#10;[server] State    :W  :server shows error state of HwControl class&#13;&#10;   DiasMaster   :W  :server which is connected to DiasMaster&#13;&#10;[members] s_DiasMaster  :W  :pointer to DiasMaster functions and settings&#13;&#10;" Name="DiasMaster.Write"/>
	FUNCTION VIRTUAL GLOBAL DiasMaster::Write
		VAR_INPUT
			input (EAX) 	: DINT;
		END_VAR
		VAR_OUTPUT
			result (EAX) 	: DINT;
		END_VAR;

	FUNCTION VIRTUAL GLOBAL SafetyState::Read
		VAR_OUTPUT
			output (EAX) 	: DINT;
		END_VAR;
  //Tables:
	FUNCTION @STD
		VAR_OUTPUT
			ret_code	: CONFSTATES;
		END_VAR;
	FUNCTION GLOBAL TAB @CT_;
END_CLASS;

#pragma using HwcLogging
#pragma using HWRtPostScan
#pragma using SafetyManager

#pragma usingLtd VaranManager

#pragma using VaranManager_Base
#pragma using VaranManager

#include <lsl_st_xtimer.h>

(************************************************************************************
*
*	Class controlls timing of DiasMaster and VaranMaster (later for more VaranMasters)
*	Created : Sigmatek	/	SR	/	March-April 2006
*	Changes :
*
*
*   FOR NEWER CHANGES SEE REVISION DOCUMENTATION OF CLASS
*
*
*		1.3 => 1.4 	/   30.06.2008
*           - [DB 884]: prevent exception in method DiasMaster::Write
*		1.2 => 1.3  /   21.03.2008
*			- [DB 817]: set RtDebug-Flag in DiasMaster
*		1.1 => 1.2	/	29.02.2008
*			- [DB 770]:	add function to get Rt-Debug State
*		1.0 => 1.1	/	28.11.2006
*			first library version
*		0.2 => 1.0	/	09.10.2006
*			initial version
*		0.1 => 0.2	/	13.06.2006
*			second testversion
*		0.0	=> 0.1	/	10.04.2006
*			first testversion for fair in Hannover
*
************************************************************************************)
VAR_PRIVATE
  HwControlThis             : ^void;
  bPostInitFinished         : BOOL;
END_VAR

#ifdef DiasMasterC_Profiler
  VAR_GLOBAL

    HWC_Time_RTPostscan		: STRUCT
        _min 	: udint;
        _max 	: udint;
        avg 	: udint;
        run 	: udint;
        sum 	: udint;
        start : udint;
        stop 	: udint;
        diff 	: udint;
        init	: udint;
        initfl: bool;

    END_STRUCT;
  END_VAR
#endif

//Has to be activated in HwControl.h
#ifdef HWCONTROL_TIME_MEASUREMENT
  #pragma message("***************************************")
  #pragma message("HWCONTROL_TIME_MEASUREMENT is activated")
  #pragma message("***************************************")
#endif

// Method define because we need poiner to method
FUNCTION GLOBAL LDR_InstallPostInitCB
  VAR_INPUT
    pThis       : ^VirtualBase;
    pCmdSvr     : ^SVRCHCMD;
    newInstCmd  : UINT;
  END_VAR;

FUNCTION HwControl::HwControl
  VAR_OUTPUT
    ret_code 	: ConfStates;
  END_VAR
  VAR
    i : USINT;
  END_VAR

  //Set supported features of HwControl (only for compatibility reasons)
  SupportedFeatures.PostInitDoneCmdCalled := TRUE;  //Flag which indicates, that the PostinitDone CMD will be called in PostInit for every logged in class
  SupportedFeatures.CalculateTaskInfo     := TRUE;  //Flag which indicates, that the HwControl calculate the task settings (RT,CY) for each core due to the logged in objects

  //Initialize us_CoreSelect
  for i:= 0 to TASK_SELECT_COREMAX do
    aTaskInfoCore[i].us_CoreSelect := i;
  end_for;

  //Store this pointer of HwControl
  HwControlThis := this;

  HWC_LogInit();

#ifdef HWC_ENABLE_SPAM_PROTECTION
  // pause spam protection to allow complete logging during init and post init phase
  HwcLogging.OverrideSpamProtection.Write(input:=1);
#endif

  //Initialize in constructor to be sure that flag is false also in the complete init phase
  bPostInitFinished := FALSE;

  ret_code := C_OK;

END_FUNCTION

FUNCTION VIRTUAL GLOBAL HwControl::Init
  VAR
    MyPara          : CmdStruct;
    MyResult        : results;
    udFirstCallCnt  : UDINT;
    pHelp           : ^t_HwObjectListCallFirst;
    retcode         : DINT;
#ifdef HWCONTROL_TIME_MEASUREMENT
    i : USINT;
#endif
  END_VAR

  //-------------------------------------------------------------------------------------------------------------
  //First Init - phase
  if ( us_InitCounter = 0 ) then

    //set this pointer to Rt-Debug function
    if ( OS_CILGet( "DEBUGAPI", #p_DebugAPI ) = SYS_ERR_NONE ) then

      //look if realtime debug option is used (our Rt-task is running even if realtime of user is debugged)
      RtDebug := RtDebug.read();

    end_if;

     //get cil interface to trigger watchdog
    OS_CILGet( INTERFACE_WATCHDOG, #p_WatchdogAPI );

    //Get OS-Interface for system info (To get amount of CPU Cores)
    if OS_CILGET(INTERFACE_LSL_SYSINFO, #pLSLSysInfo) <> SYS_ERR_NONE then
      pLSLSysInfo := NIL;
      ud_CPUCoreCount := 1; //Standard
    else
      retcode$DINT := OS_SYSINFO_GET_PROP(pLSLSysInfo, LSL_SYSINFO_ID_CPU_COUNT, #ud_CPUCoreCount, sizeof(ud_CPUCoreCount));

      if retcode <> LSL_SYSINFO_ERR_NONE then
        ud_CPUCoreCount := 1; //Standard
      end_if;
    end_if;

    //Get information if the use of the additional cores for Realtime and Cyclic is enabled

    //_Firstscan ... (*AT % M 0EB8*), _cpus_RtCyEnabled ... (*AT % M 0F21*)
    //Offset between these variables is 16#69

    //Use pointer instead of the name to be compatible with old Loader versions (old loader does not have this variable --> compiler error)
    us_CPUsRtCyEnabled := ( ( #_Firstscan + 16#69 )$^USINT)^; //0... information not available, x ... number of core with enabled RT/CY threads

  end_if;

  //-------------------------------------------------------------------------------------------------------------
  //in last init phase we call DiasMaster init functions, bring our realtime task to first position and start it
  if ( _Firstscan = TRUE ) then

    // tell the loader that we need a post init phase
    if InstallPostInitCB() <> 0 then
      HWC_LogError(this, "@014F (HwControl::Init) Failed to install post init callback!");
    end_if;

    //look if DiasMaster is also used
    if ( s_DiasMaster.p_Functions <> NIL ) then
      //make some initialization in DiasMaster before we can start our realtime task
      CallPtr	( p_function	:= s_DiasMaster.p_Functions^.p_FinishIMProg
              , p_this		  := s_DiasMaster.p_Functions^.p_This
              );
    end_if;

    // if there is no post init => we have to start the realtime from here
    if b_PostInitInstalled = FALSE then
      // Call own NewInst with CMD_POST_INIT_CALL. For sorting VaranDOs, starting RT task, init diasmaster")
      MyPara.uiCmd := CMD_POST_INIT_CALL;
      Control.NewInst(pPara:=#MyPara, pResult:=#MyResult);
    end_if;

    // if there is no varan manager and no diasmaster => we have to trigger the CDIAS watchdog for internal IOs (ETV Edge)
    if (VaranManagersAvailable = 0) & (s_DiasMaster.p_Functions = NIL) then
      OS_CILGET( "CDIASWATCHDOG", #pSCDW );
    end_if;

#ifdef HWCONTROL_TIME_MEASUREMENT
    OS_CILGet("SYSTRACE", #pSystrace$void);

    //AddTraceKeyVal is only supported with RTK and Salamander with the new kernel ( >= 9.3.0)
    //This function is supported for the CP731 but has caused problems with another PLC (WA042).
    //Therefore this feature has been deactivated for versions 09.02.xxx.
      if ( _RtOSVersion < 16#9100 ) | ( _RtOSversion >= 0x9300 ) then

      //Add Trace key values for a better visualisation in trace view
      OS_AddTraceKeyVal(pSystrace, TRECGRP_USER0, HWCONTROL_SYSTRACE_RTPRESCAN_START,                    "HwControl - Prescan: Start Realtime");
      OS_AddTraceKeyVal(pSystrace, TRECGRP_USER0, HWCONTROL_SYSTRACE_RTPRESCAN_START_FIRST_CALL_OBJECTS, "HwControl - Prescan: Start First Call Objects");
      OS_AddTraceKeyVal(pSystrace, TRECGRP_USER0, HWCONTROL_SYSTRACE_RTPRESCAN_START_VARAN_MANAGERS,     "HwControl - Prescan: Start VARAN Manager");
      OS_AddTraceKeyVal(pSystrace, TRECGRP_USER0, HWCONTROL_SYSTRACE_RTPRESCAN_START_HW_OBJECTS,         "HwControl - Prescan: Start HW Objects (SDIAS,IOs)");
      OS_AddTraceKeyVal(pSystrace, TRECGRP_USER0, HWCONTROL_SYSTRACE_RTPRESCAN_START_DIAS_CDIAS_OTHER,   "HwControl - Prescan: Start other Objects (DIAS,SpecialHW)");
      OS_AddTraceKeyVal(pSystrace, TRECGRP_USER0, HWCONTROL_SYSTRACE_RTPRESCAN_FINISH,                   "HwControl - Prescan: Finished RtWork");

      OS_AddTraceKeyVal(pSystrace, TRECGRP_USER0, HWCONTROL_SYSTRACE_RTPOSTSCAN_START,                   "HwControl - Postscan: Start Postscan");
      OS_AddTraceKeyVal(pSystrace, TRECGRP_USER0, HWCONTROL_SYSTRACE_RTPOSTSCAN_START_VARAN_MANAGERS,    "HwControl - Postscan: Start VARAN Manager");
      OS_AddTraceKeyVal(pSystrace, TRECGRP_USER0, HWCONTROL_SYSTRACE_RTPOSTSCAN_START_HW_OBJECTS,        "HwControl - Postscan: Start HW Objects (SDIAS,IOs):");
      OS_AddTraceKeyVal(pSystrace, TRECGRP_USER0, HWCONTROL_SYSTRACE_RTPOSTSCAN_FINISH,                  "HwControl - Postscan: Finished RtPostScan");

      OS_AddTraceKeyVal(pSystrace, TRECGRP_USER0, HWCONTROL_SYSTRACE_CYWORK_START,                       "HwControl - Cywork: Start Cywork");
      OS_AddTraceKeyVal(pSystrace, TRECGRP_USER0, HWCONTROL_SYSTRACE_CYWORK_START_VARAN_MANAGERS,        "HwControl - Cywork: Start VARAN Manager");
      OS_AddTraceKeyVal(pSystrace, TRECGRP_USER0, HWCONTROL_SYSTRACE_CYWORK_START_HW_OBJECTS,            "HwControl - Cywork: Start HW Objects (SDIAS,IOs)");
      OS_AddTraceKeyVal(pSystrace, TRECGRP_USER0, HWCONTROL_SYSTRACE_CYWORK_FINISH,                      "HwControl - Cywork: Finished Cywork");

    end_if;

    //Initialize min values of time measurement
    for i:= 0 to TASK_SELECT_COREMAX-1 do

      aHwControl_Times[i].sRtPrescan_Total.MinTime          := 16#FFFF;
      aHwControl_Times[i].sRtPrescan_FirstCallHW.MinTime    := 16#FFFF;
      aHwControl_Times[i].sRtPrescan_HwObjects.MinTime      := 16#FFFF;
      aHwControl_Times[i].sRtPrescan_Varan.MinTime          := 16#FFFF;
      aHwControl_Times[i].sRtPrescan_Other.MinTime          := 16#FFFF;

      aHwControl_Times[i].sRtPostscan_Total.MinTime         := 16#FFFF;
      aHwControl_Times[i].sRtPostscan_HwObjects.MinTime     := 16#FFFF;
      aHwControl_Times[i].sRtPostscan_Varan.MinTime         := 16#FFFF;

      aHwControl_Times[i].sCyWork_Total.MinTime             := 16#FFFF;
      aHwControl_Times[i].sCyWork_HwObjects.MinTime         := 16#FFFF;
      aHwControl_Times[i].sCyWork_Varan.MinTime             := 16#FFFF;

    end_for;

#endif

    // if first call objects logged in arrange them to a daisy chain
    if bCallFirstObjects then
      OS_CILGet("SYSTRACE", #pSystrace$void);

      //AddTraceKeyVal is only supported with RTK and Salamander with the new kernel ( >= 9.3.0)
      if ( _RtOSVersion < 16#9100 ) | ( _RtOSversion >= 0x9300 ) then
        OS_AddTraceKeyVal(pSystrace, TRECGRP_USER0, HWCONTROL_SYSTRACE_RTPRESCAN_FINISHED_FIRST_CALL_OBJECTS, "HwControl - Prescan: Finished Call of First Call Objects");
      end_if;

      bCallFirstObjects := FALSE;
      for udFirstCallCnt := 0 to HWCONTROL_MAX_FIRSTCALL_OBJECTS-1 do
        if sCallFirstObjects[udFirstCallCnt].pThis <> NIL then
          if bCallFirstObjects = FALSE then
            pCallFirstObjects$pVoid := To_StdLib.Malloc(size:=sizeof(t_HwObjectListCallFirst));
            pHelp                   := pCallFirstObjects;
            bCallFirstObjects       := TRUE;
          else
            pHelp^.pNext$pVoid      := To_StdLib.Malloc(size:=sizeof(t_HwObjectListCallFirst));
            pHelp                   := pHelp^.pNext;
          end_if;
          pHelp^.pThis              := sCallFirstObjects[udFirstCallCnt].pThis;
          pHelp^.udLoggedInNumber   := udFirstCallCnt;
          pHelp^.us_CoreSelect      := sCallFirstObjects[udFirstCallCnt].us_CoreSelect;
          pHelp^.ud_RtTime_us       := sCallFirstObjects[udFirstCallCnt].ud_RtTime_us;
          pHelp^.ud_CyTime_us       := sCallFirstObjects[udFirstCallCnt].ud_CyTime_us;
          pHelp^.pNext              := NIL;
        end_if;
      end_for;
      bCallFirstObjects := TRUE;
    end_if;
  end_if;

  us_InitCounter += 1;		//increment init phase counter

//-------------------------------------Profiler Start----------------------------------------------
  //#WP001 start
  #ifdef DiasMasterC_Profiler
    HWC_Time_RTPostscan.sum 	:= 0;
    HWC_Time_RTPostscan.run 	:= 0;
    HWC_Time_RTPostscan._max 	:= 0;
    HWC_Time_RTPostscan._min 	:= 16#ffffffff;
    HWC_Time_RTPostscan.init  := OS_readmicrosec();
  #endif
  //#WP001 end
//-------------------------------------Profiler End------------------------------------------------

END_FUNCTION //VIRTUAL GLOBAL HwControl::Init

FUNCTION VIRTUAL GLOBAL HwControl::RtWork
  VAR_INPUT
    EAX 	: UDINT;
  END_VAR
  VAR_OUTPUT
    state (EAX) 	: UDINT;
  END_VAR
  VAR
    us_CoreSelect : USINT;
    pHelp         : ^t_HwObjectListElement;
    udOldCnt      : UDINT;
#ifdef HWCONTROL_TIME_MEASUREMENT
    udTimeMeasure1 : UDINT;
    udTimeMeasure2 : UDINT;
#endif
  END_VAR

  us_CoreSelect := TASK_SELECT_CORE0;

#ifdef HWCONTROL_TIME_MEASUREMENT
  OS_MakeTraceEntry(pSystrace, HWCONTROL_SYSTRACE_TYPE, HWCONTROL_SYSTRACE_RTPRESCAN_START,us_CoreSelect);
#endif

  //if class is ok
  if ( HwControl::State = _ClassOk ) then

    // if interface is available trigger watchdog
    //**********************************************************************************************************************************************************
    if p_WatchdogAPI then
      OS_WD_TRIGGER(p_WatchdogAPI);

    // trigger watchdog (pointer only valid if no varan manager and diasmaster available)
    elsif pSCDW then
      SCDW_CDWTRIGGER();
    end_if;

    // special classes with first call priority, which are controlled by HwControl
    //**********************************************************************************************************************************************************
#ifdef HWCONTROL_TIME_MEASUREMENT
    OS_MakeTraceEntry(pSystrace, HWCONTROL_SYSTRACE_TYPE, HWCONTROL_SYSTRACE_RTPRESCAN_START_FIRST_CALL_OBJECTS,us_CoreSelect);
    udTimeMeasure1 := OS_READMICROSEC();
#endif

    UpdateRtFirstCallObjects(us_CoreSelect);

#ifdef HWCONTROL_TIME_MEASUREMENT
    udTimeMeasure2 := OS_READMICROSEC();
    aHwControl_Times[us_CoreSelect].sRtPrescan_FirstCallHW.ActTime := udTimeMeasure2 - udTimeMeasure1;
#endif

    //Increment timestamp for SmartIO modules
    aTaskInfoCore[us_CoreSelect].uiHwTimeStamp_us += (aTaskInfoCore[us_CoreSelect].ud_MyRtTaskTime_us)$UINT;

    //Send Sync for DiasMaster
    //**********************************************************************************************************************************************************
    if ( s_DiasMaster.p_Functions <> NIL ) then
      //if call time for dias master is reached
      if ( s_DiasMaster.ud_Counter = s_DiasMaster.p_Functions^.ud_DiasTime ) then

        CallPtr	( p_function	:= s_DiasMaster.p_Functions^.p_SendSync
                , p_this		  := s_DiasMaster.p_Functions^.p_This
                );
      end_if;
    end_if;

    //Update Realtime of all varanmanagers which are running on core 0
    //**********************************************************************************************************************************************************
#ifdef HWCONTROL_TIME_MEASUREMENT
    OS_MakeTraceEntry(pSystrace, HWCONTROL_SYSTRACE_TYPE, HWCONTROL_SYSTRACE_RTPRESCAN_START_VARAN_MANAGERS,us_CoreSelect);
    udTimeMeasure1 := OS_READMICROSEC();
#endif

    UpdateRtVaranManager(us_CoreSelect);

#ifdef HWCONTROL_TIME_MEASUREMENT
    udTimeMeasure2 := OS_READMICROSEC();
    aHwControl_Times[us_CoreSelect].sRtPrescan_Varan.ActTime := udTimeMeasure2 - udTimeMeasure1;
#endif

    //DiasMaster Call Rt
    //**********************************************************************************************************************************************************
#ifdef HWCONTROL_TIME_MEASUREMENT
    OS_MakeTraceEntry(pSystrace, HWCONTROL_SYSTRACE_TYPE, HWCONTROL_SYSTRACE_RTPRESCAN_START_DIAS_CDIAS_OTHER,us_CoreSelect);
    udTimeMeasure1 := OS_READMICROSEC();
#endif

    //Only call DIAS from core 0
    if ( s_DiasMaster.p_Functions <> NIL ) then
      //if call time for dias master is reached
      if ( s_DiasMaster.ud_Counter = s_DiasMaster.p_Functions^.ud_DiasTime ) then

        //set task time counter to HwControl task time
        s_DiasMaster.ud_Counter := aTaskInfoCore[us_CoreSelect].ud_MyRtTaskTime_us;

        CallPtr	( p_function	:= s_DiasMaster.p_Functions^.p_RtFunction
                , p_this		  := s_DiasMaster.p_Functions^.p_This
                );

      else
        //add task time to counter
        s_DiasMaster.ud_Counter += aTaskInfoCore[us_CoreSelect].ud_MyRtTaskTime_us;
      end_if;
    end_if;

    // special classes, which are controlled by HwControl (Modules which are added via AddSpecialHW)
    if pSpecialObjects then
      pHelp := pSpecialObjects;
      while pHelp <> NIL do
        pHelp^.pThis^.RtWork(0);
        pHelp := pHelp^.pNext;
      end_while;
    end_if;

#ifdef HWCONTROL_TIME_MEASUREMENT
    udTimeMeasure2 := OS_READMICROSEC();
    aHwControl_Times[us_CoreSelect].sRtPrescan_Other.ActTime := udTimeMeasure2 - udTimeMeasure1;
#endif

    // objects, which are controlled by HwControl
    //**********************************************************************************************************************************************************
#ifdef HWCONTROL_TIME_MEASUREMENT
    OS_MakeTraceEntry(pSystrace, HWCONTROL_SYSTRACE_TYPE, HWCONTROL_SYSTRACE_RTPRESCAN_START_HW_OBJECTS,us_CoreSelect);
    udTimeMeasure1 := OS_READMICROSEC();
#endif

    UpdateRtLoginObjects(usCoreSelect:= us_CoreSelect);

#ifdef HWCONTROL_TIME_MEASUREMENT
    udTimeMeasure2 := OS_READMICROSEC();
    aHwControl_Times[us_CoreSelect].sRtPrescan_HwObjects.ActTime := udTimeMeasure2 - udTimeMeasure1;
#endif

    // if someone wants to debug realtime or we are in startup phase (only 1 rt object possible to start while init is running)
    //**********************************************************************************************************************************************************
    if RtDebug | (_FirstScan & (aTaskInfoCore[us_CoreSelect].b_PostScanStarted = FALSE)) then
      PostScanWork(us_CoreSelect);
      if (RtDebug = 0) then
        aTaskInfoCore[us_CoreSelect].ud_LastPostScanWorkCall := OS_READMICROSEC();
      end_if;
    else
      //check for active realtime synchronisation
      if sRtTaskControl.b_RtTaskControlActive = TRUE then

        //increment finished counter for this rt prescan - counter is decrement after syncronizing
        udOldCnt := sigclib_atomic_incU32(pValue:=#sRtTaskControl.udPreRtCnt);

        //if old counter is all cores -1 then is the last prescan rt reached
        if udOldCnt >= sRtTaskControl.usCoresRtActive - 1 then

          //all rt tasks are finished -> free mutex
          OS_MT_SIGNAL(sRtTaskControl.pvPreRtSyncTaskEvent);

          sigclib_atomic_decU32(pValue:=#sRtTaskControl.udPreRtCnt);

          //if the counter reached zero we know all other PreScans at Wait State are unlocked again
          while sigclib_atomic_getU32(pValue:=#sRtTaskControl.udPreRtCnt) <> 0 do

          end_while;

          //reset PreScan mutex
          OS_MT_RESETEVENT(sRtTaskControl.pvPreRtSyncTaskEvent);
        else
          //wait for other rt task to be finished
          OS_MT_WAIT(sRtTaskControl.pvPreRtSyncTaskEvent);
          sigclib_atomic_decU32(pValue:=#sRtTaskControl.udPreRtCnt);
        end_if;
      end_if;
    end_if;
  end_if;

#ifdef HWCONTROL_TIME_MEASUREMENT
  OS_MakeTraceEntry(pSystrace, HWCONTROL_SYSTRACE_TYPE, HWCONTROL_SYSTRACE_RTPRESCAN_FINISH,us_CoreSelect);
  CalcTimeMeasurementPreScan(#aHwControl_Times[us_CoreSelect]);
#endif

  state := READY;

END_FUNCTION

FUNCTION HwControl::RtPreScan_CoreX
  VAR_INPUT
    pCoreSelect 	: ^void;
  END_VAR
  VAR
    us_CoreSelect : USINT;
    udOldCnt : UDINT;
#ifdef HWCONTROL_TIME_MEASUREMENT
    udTimeMeasure1 : UDINT;
    udTimeMeasure2 : UDINT;
#endif
  END_VAR

  this := HwControlThis$^HWControl;
  us_CoreSelect := pCoreSelect^$USINT;

#ifdef HWCONTROL_TIME_MEASUREMENT
  OS_MakeTraceEntry(pSystrace, HWCONTROL_SYSTRACE_TYPE, HWCONTROL_SYSTRACE_RTPRESCAN_START,us_CoreSelect);
  udTimeMeasure1 := OS_READMICROSEC();
#endif

  //if class is ok
  if ( HwControl::State = _ClassOk ) then

    // special classes with first call priority, which are controlled by HwControl
    //**********************************************************************************************************************************************************
#ifdef HWCONTROL_TIME_MEASUREMENT
    OS_MakeTraceEntry(pSystrace, HWCONTROL_SYSTRACE_TYPE, HWCONTROL_SYSTRACE_RTPRESCAN_START_FIRST_CALL_OBJECTS,us_CoreSelect);
    udTimeMeasure1 := OS_READMICROSEC();
#endif

    UpdateRtFirstCallObjects(us_CoreSelect);

#ifdef HWCONTROL_TIME_MEASUREMENT
    udTimeMeasure2 := OS_READMICROSEC();
    aHwControl_Times[us_CoreSelect].sRtPrescan_FirstCallHW.ActTime := udTimeMeasure2 - udTimeMeasure1;
#endif

    aTaskInfoCore[us_CoreSelect].uiHwTimeStamp_us += (aTaskInfoCore[us_CoreSelect].ud_MyRtTaskTime_us)$UINT;

    //Update Realtime of all varanmanagers which are running on core 0
    //**********************************************************************************************************************************************************
#ifdef HWCONTROL_TIME_MEASUREMENT
    OS_MakeTraceEntry(pSystrace, HWCONTROL_SYSTRACE_TYPE, HWCONTROL_SYSTRACE_RTPRESCAN_START_VARAN_MANAGERS,us_CoreSelect);
    udTimeMeasure1 := OS_READMICROSEC();
#endif

    UpdateRtVaranManager(us_CoreSelect);

#ifdef HWCONTROL_TIME_MEASUREMENT
    udTimeMeasure2 := OS_READMICROSEC();
    aHwControl_Times[us_CoreSelect].sRtPrescan_Varan.ActTime := udTimeMeasure2 - udTimeMeasure1;
#endif

    // objects, which are controlled by HwControl
    //**********************************************************************************************************************************************************
#ifdef HWCONTROL_TIME_MEASUREMENT
    OS_MakeTraceEntry(pSystrace, HWCONTROL_SYSTRACE_TYPE, HWCONTROL_SYSTRACE_RTPRESCAN_START_HW_OBJECTS,us_CoreSelect);
    udTimeMeasure1 := OS_READMICROSEC();
#endif

    UpdateRtLoginObjects(usCoreSelect:= us_CoreSelect);

#ifdef HWCONTROL_TIME_MEASUREMENT
    udTimeMeasure2 := OS_READMICROSEC();
    aHwControl_Times[us_CoreSelect].sRtPrescan_HwObjects.ActTime := udTimeMeasure2 - udTimeMeasure1;
#endif

    // if someone wants to debug realtime or we are in startup phase (only 1 rt object possible to start while init is running)
    //**********************************************************************************************************************************************************
    if RtDebug | (_FirstScan & (aTaskInfoCore[us_CoreSelect].b_PostScanStarted = FALSE)) then
      PostScanWork(us_CoreSelect);
      if (RtDebug = 0) then
        aTaskInfoCore[us_CoreSelect].ud_LastPostScanWorkCall := OS_READMICROSEC();
      end_if;
    else
      //check for active realtime synchronisation
      if sRtTaskControl.b_RtTaskControlActive = TRUE then

        //increment finished counter for this rt prescan - counter is decrement after syncronizing
        udOldCnt := sigclib_atomic_incU32(pValue:=#sRtTaskControl.udPreRtCnt);

        //if old counter is all cores -1 then is the last prescan rt reached
        if udOldCnt >= sRtTaskControl.usCoresRtActive - 1 then

          //all rt tasks are finished -> free mutex
          OS_MT_SIGNAL(sRtTaskControl.pvPreRtSyncTaskEvent);

          sigclib_atomic_decU32(pValue:=#sRtTaskControl.udPreRtCnt);

          //if the counter reached zero we know all other PreScans at Wait State are unlocked again
          while sigclib_atomic_getU32(pValue:=#sRtTaskControl.udPreRtCnt) <> 0 do

          end_while;
          //reset PreScan mutex
          OS_MT_RESETEVENT(sRtTaskControl.pvPreRtSyncTaskEvent);
        else
          //wait for other rt task to be finished
          OS_MT_WAIT(sRtTaskControl.pvPreRtSyncTaskEvent);
          sigclib_atomic_decU32(pValue:=#sRtTaskControl.udPreRtCnt);
        end_if;
      end_if;
    end_if;
  end_if;

#ifdef HWCONTROL_TIME_MEASUREMENT
  OS_MakeTraceEntry(pSystrace, HWCONTROL_SYSTRACE_TYPE, HWCONTROL_SYSTRACE_RTPRESCAN_FINISH,us_CoreSelect);
  CalcTimeMeasurementPreScan(#aHwControl_Times[us_CoreSelect]);
#endif

END_FUNCTION

FUNCTION HwControl::RtPostScan_CoreX
  VAR_INPUT
    pCoreSelect 	: ^void;
  END_VAR
  VAR
    us_CoreSelect : USINT;
    udOldCnt : UDINT;
  END_VAR

  this := HwControlThis$^HWControl;
  us_CoreSelect := pCoreSelect^$USINT;

  if sRtTaskControl.b_RtTaskControlActive = TRUE then

    //increment PostScan start counter for this rt PostScan - counter is decrement after syncronizing
    udOldCnt := sigclib_atomic_incU32(pValue:=#sRtTaskControl.udPostRtCnt);

    //if old counter is all cores -1 then is the last postscan rt reached
    if udOldCnt >= sRtTaskControl.usCoresRtActive - 1 then

      //all PostScans tasks are reached -> free mutex
      OS_MT_SIGNAL(sRtTaskControl.pvPostRtSyncTaskEvent);

      sigclib_atomic_decU32(pValue:=#sRtTaskControl.udPostRtCnt);

      //if the counter reached zero we know all other PostScans at Wait State are unlocked again
      while sigclib_atomic_getU32(pValue:=#sRtTaskControl.udPostRtCnt) <> 0 do

      end_while;

      //reset PreScan mutex
      OS_MT_RESETEVENT(sRtTaskControl.pvPostRtSyncTaskEvent);
    else
      //wait for other rt task to be finished
      OS_MT_WAIT(sRtTaskControl.pvPostRtSyncTaskEvent);
      sigclib_atomic_decU32(pValue:=#sRtTaskControl.udPostRtCnt);
    end_if;
  end_if;

  // first time postscan is called by os
  if aTaskInfoCore[us_CoreSelect].b_PostScanStarted = FALSE then
    aTaskInfoCore[us_CoreSelect].b_PostScanStarted := TRUE;
    if p_WatchdogAPI then
      //turn of watchdogtask of os because we trigger it in application
      OS_WD_SETPROPERTY(p_WatchdogAPI, Property:=WD_PROP_APPL_WD, value:=1); // 1 to disable autotrigger
    end_if;
    // if we've already done postscan work from prescan, don't do anything here
    aTaskInfoCore[us_CoreSelect].ud_FirstPostScanCall := OS_READMICROSEC();
    // check if already called in same cycle => my task time in ns recalculated to 80 percent of the task time in µs
    if (aTaskInfoCore[us_CoreSelect].ud_FirstPostScanCall - aTaskInfoCore[us_CoreSelect].ud_LastPostScanWorkCall) < ((aTaskInfoCore[us_CoreSelect].ud_MyRtTaskTime_us * 80) / 100) then
      return;
    end_if;
  end_if;

  PostScanWork(us_CoreSelect);

END_FUNCTION

FUNCTION HwControl::CyWork_CoreX
  VAR_INPUT
    pCoreSelect 	: ^void;
  END_VAR
  VAR
    us_CoreSelect : USINT;
    pHelp         : ^t_HwObjectListElement;
    pOneManager   : ^t_OneVaranManager;
    i             : USINT;
#ifdef HWCONTROL_TIME_MEASUREMENT
    udTimeMeasure1 : UDINT;
    udTimeMeasure2 : UDINT;
#endif
  END_VAR

  this := HwControlThis$^HWControl;

  us_CoreSelect := pCoreSelect^$USINT;

#ifdef HWCONTROL_TIME_MEASUREMENT
  OS_MakeTraceEntry(pSystrace, HWCONTROL_SYSTRACE_TYPE, HWCONTROL_SYSTRACE_CYWORK_START,us_CoreSelect);
#endif

  //Update cyclic of all varanmanagers
  //*****************************************************************************
#ifdef HWCONTROL_TIME_MEASUREMENT
  udTimeMeasure1 := OS_READMICROSEC();
  OS_MakeTraceEntry(pSystrace, HWCONTROL_SYSTRACE_TYPE, HWCONTROL_SYSTRACE_CYWORK_START_VARAN_MANAGERS,us_CoreSelect);
#endif

  pOneManager := #a_VaranManager[0];
  for i := 0 TO (MAX_VARAN_MANAGERS - 1) do
    //Look for right core
    if pOneManager^.us_CoreSelect = us_CoreSelect then

      //Check for valid manager
      if pOneManager^.p_Functions <> NIL  then

        //Only call cywork if it is time to call it
        if pOneManager^.ud_CounterCy = pOneManager^.ud_CyTime_us then
          pOneManager^.ud_CounterCy := 0;
          pOneManager^.p_Functions^.p_This^.CyWork();
        end_if;

        pOneManager^.ud_CounterCy += aTaskInfoCore[us_CoreSelect].ud_MyCyTaskTime_us;

      end_if;
    end_if;
    pOneManager += SIZEOF(t_OneVaranManager);
  end_for;

#ifdef HWCONTROL_TIME_MEASUREMENT
  udTimeMeasure2 := OS_READMICROSEC();
  aHwControl_Times[us_CoreSelect].sCyWork_Varan.ActTime := udTimeMeasure2 - udTimeMeasure1;
#endif

  //Update cyclic of other objects
  //*****************************************************************************
#ifdef HWCONTROL_TIME_MEASUREMENT
  OS_MakeTraceEntry(pSystrace, HWCONTROL_SYSTRACE_TYPE, HWCONTROL_SYSTRACE_CyWORK_START_HW_OBJECTS,us_CoreSelect);
  udTimeMeasure1 := OS_READMICROSEC();
#endif

  if pHwControlLogins then
    pHelp := pHwControlLogins;
    while pHelp <> NIL do
      if pHelp^.bdSettings.Cyclic & pHelp^.us_CoreSelect = us_CoreSelect then
        pHelp^.pThis^.CyWork(0);
      end_if;
      pHelp := pHelp^.pNext;
    end_while;
  end_if;

#ifdef HWCONTROL_TIME_MEASUREMENT
  udTimeMeasure2 := OS_READMICROSEC();
  aHwControl_Times[us_CoreSelect].sCyWork_HwObjects.ActTime := udTimeMeasure2 - udTimeMeasure1;

  OS_MakeTraceEntry(pSystrace, HWCONTROL_SYSTRACE_TYPE, HWCONTROL_SYSTRACE_CYWORK_FINISH,us_CoreSelect);
  CalcTimeMeasurementCyclic(#aHwControl_Times[us_CoreSelect]);
#endif

END_FUNCTION

FUNCTION GLOBAL HwControl::AddVaranManager
  VAR_INPUT
    ud_manager_number 	: UDINT;
    p_function_list 	  : ^void;
    us_CoreSelect 	    : USINT;(* := 0 *)
    ud_RtTime_us 	      : UDINT;(* := 0 *)
    ud_CyTime_us 	      : UDINT;(* := 0 *)
  END_VAR
  VAR_OUTPUT
    sd_retval 	: DINT;
  END_VAR

  // is class ok
  if ( State = _ClassOk ) then

    //Check if selected core is available at this CPU
    if ( us_CoreSelect > TASK_SELECT_CORE0 ) & (us_CoreSelect > (ud_CPUCoreCount-1)) then
      sd_retval := -4;    //Invalid Core selected
      HWC_LogValue2(this,"@0150 (HwControl::AddVaranManager) Invalid parameter us_CoreSelect 0x{0}. CPU only has 0x{1} core(s)", us_CoreSelect, ud_CPUCoreCount);
      return;

    //Check if the use of the additional cores for Realtime and Cyclic is enabled
    elsif ( us_CoreSelect > TASK_SELECT_CORE0 ) & (us_CoreSelect > (us_CPUsRtCyEnabled-1)) then
      sd_retval := 11;
      HWC_LogError(this, "@0151 (HwControl::AddVaranManager) Rt/Cy Tasks are not enabled for the additional cores. Please use <SET MULTICOREOBJS 1> in autoexec.lsl");
      return;

    //Check if the LSL_I_TASK Interface version supports multicore
    elsif ( us_CoreSelect > TASK_SELECT_CORE0 ) & ( Get_ITASK_Version() < LSL_ITASK_VERSION_MULTICORE_SUPPORT ) then
      sd_retval := -5;
      HWC_LogError(this, "@0152 (HwControl::AddVaranManager) Invalid CPU-Core selected for this CPU. Version of LSL_ITASK Interface doesn't support multicore");
      return;

    //Check if coreselect is supported by HwControl already
    elsif ( us_CoreSelect > TASK_SELECT_COREMAX ) then
      sd_retval := -6; //Failed to install realtime task
      HWC_LogValue2(this, "@0153 (HwControl::AddVaranManager) Invalid parameter us_CoreSelect 0x{0}. Max. us_CoreSelect by HwControl is 0x{1}",us_CoreSelect,TASK_SELECT_COREMAX);
      return;
    end_if;

    //Check if Rt time is smaller than maintimer
    if ( ud_RtTime_us <> 0 ) & ( ud_RtTime_us < _ClockTicks ) then
      sd_retval := -7;
      HWC_LogError(this, "@0154 (HwControl::AddVaranManager) Parameter ud_RtTime_us is smaller than CPU maintimer!");
      return;

    //Check if Rt time is not a multiple of maintimer
    elsif ( ud_RtTime_us <> 0 ) & (ud_RtTime_us MOD _ClockTicks) <> 0 then
      sd_retval := -8;
      HWC_LogError(this, "@0155 (HwControl::AddVaranManager) Parameter ud_RtTime_us not a multiple of CPU maintimer!");
      return;
    end_if;

    //Check if Cy time is smaller than maintimer
    if ( ud_CyTime_us <> 0 ) & ud_CyTime_us < _ClockTicks then
      sd_retval := -9;
      HWC_LogError(this, "@0156 (HwControl::AddVaranManager) Parameter ud_CyTime_us is smaller than CPU maintimer!");
      return;

    //Check if CY time is not a multiple of maintimer
    elsif ( ud_CyTime_us <> 0 ) & (ud_CyTime_us MOD _ClockTicks) <> 0 then
      sd_retval := -10;
      HWC_LogError(this, "@0157 (HwControl::AddVaranManager) Parameter ud_CyTime_us not a multiple of CPU maintimer!");
      return;

    end_if;

    // look if it is a correct VaranManager number
    if	(( ud_manager_number >= 0 ) &
         ( ud_manager_number <= MAX_VARAN_MANAGERS - 1 )) then

      // look if the pointer is valid
      if p_function_list then

        //is this number already in use
        if ( a_VaranManager[ ud_manager_number ].p_Functions <> NIL ) then

          State											                      := _NotInitialized;		//Set to error state
          a_VaranManager[ ud_manager_number ].p_Functions	:= NIL;
          sd_retval 										                  := -6;

          HWC_LogError(this, "@0158 (HwControl::AddVaranManager) Multiple VaranManager number!");
          return;
        end_if;

        //load pointer to varan functions
        a_VaranManager[ ud_manager_number ].p_Functions$^void := p_function_list;

        //Save core to execute task from
        a_VaranManager[ ud_manager_number ].us_CoreSelect   := us_CoreSelect;

        //set counter to time to execute task at first realtime
        if ud_RtTime_us <> 0 then
          a_VaranManager[ ud_manager_number ].ud_RtTime_us    := ud_RtTime_us;
          a_VaranManager[ ud_manager_number ].ud_CounterRt    := a_VaranManager[ ud_manager_number ].ud_RtTime_us;
        else
          a_VaranManager[ ud_manager_number ].ud_RtTime_us    := a_VaranManager[ ud_manager_number ].p_Functions^.ud_VaranTime / 1000;  //Convert from ns to µs
          a_VaranManager[ ud_manager_number ].ud_CounterRt    := a_VaranManager[ ud_manager_number ].p_Functions^.ud_VaranTime / 1000;  //Convert from ns to µs
        end_if;

        //set counter to time to execute task at first cyclic
        if ud_CyTime_us <> 0 then
          a_VaranManager[ ud_manager_number ].ud_CyTime_us    := ud_CyTime_us;
          a_VaranManager[ ud_manager_number ].ud_CounterCy    := a_VaranManager[ ud_manager_number ].ud_CyTime_us;
        else
          a_VaranManager[ ud_manager_number ].ud_CyTime_us    := a_VaranManager[ ud_manager_number ].p_Functions^.ud_VaranTime / 1000;  //Convert from ns to µs
          a_VaranManager[ ud_manager_number ].ud_CounterCy    := a_VaranManager[ ud_manager_number ].p_Functions^.ud_VaranTime / 1000;  //Convert from ns to µs
        end_if;

        sd_retval 	:= 0;

        // new varanmanager is avaliable
        VaranManagersAvailable += 1;
      else
        sd_retval := -3;			// pointer invalid
        HWC_LogError(this, "@0159 (HwControl::AddVaranManager) Invalid pointer!");
      end_if;
    else
      sd_retval := -2;			//manager number wrong
      HWC_LogError(this, "@015A (HwControl::AddVaranManager) Wrong VaranManagerNumber!");
    end_if;
  else
    sd_retval := -1; // class state not _ClassOk
    HWC_LogError(this, "@015B (HwControl::AddVaranManager) Class state is not ok!");
  end_if;

END_FUNCTION //GLOBAL HwControl::AddVaranManager

FUNCTION HwControl::CallPtr
  VAR_INPUT
    p_function	: pFct;
    p_this		  : pVoid;
  END_VAR
  VAR
    save_this   :^HwControl;
  END_VAR

  save_this := this;              // save this ptr
  this      := p_this$^HwControl; // load thispointer of object
  p_function$ObjectFunct();       // call function of object
  this      := save_this;         // restore this ptr

END_FUNCTION // HwControl::CallPtr

FUNCTION GLOBAL HwControl::GetMyTaskTime
  VAR_INPUT
    us_CoreSelect 	: DINT;(* := 0 *)
  END_VAR
  VAR_OUTPUT
    ud_task_time 	: UDINT;
  END_VAR

  //Check if we already have calculated a time for the Realtime
  ud_task_time := aTaskInfoCore[us_CoreSelect].ud_MyRtTaskTime_us * 1000;		//give back task time in ns

END_FUNCTION // HwControl::GetMyTaskTime

FUNCTION GLOBAL HwControl::SetHardwareOff
  VAR_INPUT
    e_error		: t_e_VaranErrors;
  END_VAR
  VAR
    MyPara    : CmdStruct;
    MyResult  : results;
  END_VAR

  State := e_error;

  // if a diasmaster is available => tell him
  if s_DiasMaster.p_Functions then
    MyPara.uiCmd := CMD_HWC_ERROR_TO_DIASM;
    s_DiasMaster.p_Functions^.p_This$pVirtualBase^.NewInst(#MyPara,#MyResult);
  end_if;

END_FUNCTION //GLOBAL HwControl::SetHardwareOff

FUNCTION GLOBAL HwControl::GetRtDebugState
  VAR_OUTPUT
    sd_RtDebug		: DINT;
  END_VAR

  sd_RtDebug := RtDebug.read();

END_FUNCTION //GLOBAL HwControl::GetRtDebugState

FUNCTION VIRTUAL GLOBAL HwControl::DiasMaster::Write
  VAR_INPUT
    input (EAX) 	: DINT;
  END_VAR
  VAR_OUTPUT
    result (EAX) 	: DINT;
  END_VAR

  //is it a required error from dias master?
  if input = 0 then
    State := _RequiredError;
    return;
  end_if;

  //is class ok
  if ( State = _ClassOk ) then

    s_DiasMaster.p_Functions$DINT := input;		//load pointer to DiasMaster functions

    //look if DiasMaster time is faster as the maintimer
    if ( ( s_DiasMaster.p_Functions^.ud_DiasTime ) < (_ClockTicks) ) then

      State						          := _DiasTimeError;			//Set to error state
      s_DiasMaster.p_Functions	:= NIL;
      result 						        := -1;
      HWC_LogError(this, "@015C (HwControl::DiasMaster::Write) DiasMaster time is smaller than HwControl RT-Task!");
      return;
    //look if DiasMaster time is a multiple time of our task time
    elsif ( ( s_DiasMaster.p_Functions^.ud_DiasTime ) mod (_ClockTicks) <> 0 ) then

      State						          := _DiasTimeError;			//Set to error state
      s_DiasMaster.p_Functions	:= NIL;
      result						        := -1;
      HWC_LogError(this, "@015D (HwControl::DiasMaster::Write) DiasMaster time is not a multiple of HwControl RT-Task!");
      return;
    else
      //set counter to time to execute task at first realtime
      s_DiasMaster.ud_Counter := s_DiasMaster.p_Functions^.ud_DiasTime;
      result 					    := 0;
      DiasMaster := input := 1;				//Mark server as connected right
    end_if;

    //set RtDebug-Flag for DiasMaster
    s_DiasMaster.p_Functions^.sd_RtDebug := RtDebug.Read();
  else
    result := -1;
  end_if;

END_FUNCTION

FUNCTION GLOBAL HwControl::AddSpecialHW
  VAR_INPUT
    pThis 	      : pVirtualBase;
    pRtPostScan 	: ^UDINT;
  END_VAR
  VAR_OUTPUT
    retcode 	    : DINT;
  END_VAR
  VAR
    pHelp         : ^t_HwObjectListElement;
  END_VAR

  //Attention: This function does not provide core-selection and cycle time settings (these object will be called on core 0 every time and with the calculated time)
  //If you want to use this feature please use the method AddHwObject

  if pSpecialObjects = NIL then
    pSpecialObjects$pVoid := To_StdLib.Malloc(size:=sizeof(t_HwObjectListElement));
    pHelp := pSpecialObjects;
  else
    pHelp := pSpecialObjects;
    while pHelp^.pNext <> NIL do
      pHelp := pHelp^.pNext;
    end_while;
    pHelp^.pNext$pVoid := To_StdLib.Malloc(size:=sizeof(t_HwObjectListElement));
    pHelp := pHelp^.pNext;
  end_if;

  if pHelp <> NIL then
    pHelp^.pThis          := pThis;
    pHelp^.bdSettings     := 0;
    pHelp^.usEscSequence  := 0;
    pHelp^.us_CoreSelect  := 0;
    pHelp^.ud_RtTime_us   := 0;
    pHelp^.ud_CyTime_us   := 0;
    pHelp^.pRtPostScan    := pRtPostScan;
    pHelp^.pNext          := NIL;

    retcode               := 0;
  else
    retcode               := -1;
  end_if;

END_FUNCTION

FUNCTION GLOBAL HwControl::AddFirstCallHW
  VAR_INPUT
    pThis 	        : pVirtualBase;
    udSelectPlace 	: UDINT;
    us_CoreSelect 	: USINT;(* := 0 *)
    ud_RtTime_us 	  : UDINT;(* := 0 *)
    ud_CyTime_us 	  : UDINT;(* := 0 *)
  END_VAR
  VAR_OUTPUT
    retcode 	: DINT;
  END_VAR

  if udSelectPlace >= HWCONTROL_MAX_FIRSTCALL_OBJECTS then
    //place is not available
    retcode := -1;
    return;
  end_if;

  if sCallFirstObjects[udSelectPlace].pThis <> NIL then
    //place is already used
    retcode := -2;
    return;
  end_if;

  if _FirstScan = TRUE then
    //object login is to late
    retcode := -3;
    return;
  end_if;

  //Check if the selected core is available on the CPU
  if ( us_CoreSelect > TASK_SELECT_CORE0 ) & (us_CoreSelect > (ud_CPUCoreCount-1)) then
    //CPU does not have the requested core
    HWC_LogValue2(this,"@0150 (HwControl::AddFirstCallHW) Invalid parameter us_CoreSelect 0x{0}. CPU only has 0x{1} core(s)", us_CoreSelect, ud_CPUCoreCount);
    retcode := -4;
    return;

  //Check if the use of the additional cores for Realtime and Cyclic is enabled
  elsif ( us_CoreSelect > TASK_SELECT_CORE0 ) & (us_CoreSelect > (us_CPUsRtCyEnabled-1)) then
    retcode := 11;
    HWC_LogError(this, "@0151 (HwControl::AddFirstCallHW) Rt/Cy Tasks are not enabled for the additional cores. Please use <SET MULTICOREOBJS 1> in autoexec.lsl");
    return;

  //Check if the LSL_I_TASK Interface version supports multicore
  elsif ( us_CoreSelect > TASK_SELECT_CORE0 ) & ( Get_ITASK_Version() < LSL_ITASK_VERSION_MULTICORE_SUPPORT ) then
    retcode := -5;
    HWC_LogError(this, "@0152 (HwControl::AddFirstCallHW) Invalid CPU-Core selected for this CPU. Version of LSL_ITASK Interface doesn't support multicore");
    return;

  //Check if coreselect is supported by HwControl already
  elsif ( us_CoreSelect > TASK_SELECT_COREMAX ) then
    retcode := -6;
    HWC_LogValue2(this, "@0153 (HwControl::AddFirstCallHW) Invalid parameter us_CoreSelect 0x{0}. Max. us_CoreSelect by HwControl is 0x{1}",us_CoreSelect,TASK_SELECT_COREMAX);
    return;
  end_if;

  //Check if Rt time is smaller than maintimer
  if ( ud_RtTime_us <> 0 ) & ( ud_RtTime_us < _ClockTicks ) then
    retcode := -7;
    HWC_LogError(this, "@0154 (HwControl::AddFirstCallHW) Parameter ud_RtTime_us is smaller than CPU maintimer !");
    return;

  //Check if Rt time is not a multiple of maintimer
  elsif ( ud_RtTime_us <> 0 ) & (ud_RtTime_us MOD _ClockTicks) <> 0 then
    retcode := -8;
    HWC_LogError(this, "@0155 (HwControl::AddFirstCallHW) Parameter ud_RtTime_us not a multiple of CPU maintimer!");
    return;
  end_if;

  //Check if Cy time is smaller than maintimer
  if ( ud_CyTime_us <> 0 ) & ud_CyTime_us < _ClockTicks then
    retcode := -9;
    HWC_LogError(this, "@0156 (HwControl::AddFirstCallHW) Parameter ud_CyTime_us is smaller than CPU maintimer !");
    return;

  //Check if CY time is not a multiple of maintimer
  elsif ( ud_CyTime_us <> 0 ) & (ud_CyTime_us MOD _ClockTicks) <> 0 then
    retcode := -10;
    HWC_LogError(this, "@0157 (HwControl::AddFirstCallHW) Parameter ud_CyTime_us not a multiple of CPU maintimer!");
    return;
  end_if;

  //set true because a first call object has logged in
  bCallFirstObjects                 := TRUE;

  //set pointer to free place
  sCallFirstObjects[udSelectPlace].pThis          := pThis;
  sCallFirstObjects[udSelectPlace].us_CoreSelect  := us_CoreSelect;
  sCallFirstObjects[udSelectPlace].ud_RtTime_us   := ud_RtTime_us;
  sCallFirstObjects[udSelectPlace].ud_CyTime_us   := ud_CyTime_us;

  //return code ok
  retcode                           := 0;

END_FUNCTION

FUNCTION GLOBAL HwControl::AddHwObject
  VAR_INPUT
    pThis 	        : pVirtualBase;
    Settings 	      : t_HwObjListSettings;
    EscapeSequence 	: USINT;(* := 0 *)
    us_CoreSelect 	: USINT;(* := 0 *)
    ud_RtTime_us 	  : UDINT;(* := 0 *)
    ud_CyTime_us 	  : UDINT;(* := 0 *)
  END_VAR
  VAR_OUTPUT
    retcode 	: DINT;
  END_VAR
  VAR
    pHelp           : ^t_HwObjectListElement;
  END_VAR

  if pThis = nil then
    //Pointer invalid
    retcode := -2;
    HWC_LogError(this,"@015E (HwControl::AddHwObject) Invalid parameter pThis.");
  end_if;

  //If Bit is false we do not take the core-select setting (maybe data is uninitialized)
  if Settings.CoreSelect = FALSE then
    us_CoreSelect := TASK_SELECT_CORE0;
  end_if;

  //If Bit is false we do not take the time settings (maybe data is uninitialized)
  if Settings.TimeSet = FALSE then
    ud_RtTime_us := 0;
    ud_CyTime_us := 0;
  end_if;

  //Check if the selected core is available on the CPU
  if ( us_CoreSelect > TASK_SELECT_CORE0 ) & (us_CoreSelect > (ud_CPUCoreCount-1)) then
    //CPU does not have the requested core
    HWC_LogValue2(this,"@0150 (HwControl::AddHwObject) Invalid parameter us_CoreSelect 0x{0}. CPU only has 0x{1} core(s)", us_CoreSelect, ud_CPUCoreCount);
    retcode := -4;
    return;

  //Check if the use of the additional cores for Realtime and Cyclic is enabled
  elsif ( us_CoreSelect > TASK_SELECT_CORE0 ) & (us_CoreSelect > (us_CPUsRtCyEnabled-1)) then
    retcode := 11;
    HWC_LogError(this, "@0151 (HwControl::AddHwObject) Rt/Cy Tasks are not enabled for the additional cores. Please use <SET MULTICOREOBJS 1> in autoexec.lsl");
    return;

  //Check if the LSL_I_TASK Interface version supports multicore
  elsif ( us_CoreSelect > TASK_SELECT_CORE0 ) & ( Get_ITASK_Version() < LSL_ITASK_VERSION_MULTICORE_SUPPORT ) then
    retcode := -5;
    HWC_LogError(this, "@0152 (HwControl::AddHwObject) Invalid CPU-Core selected for this CPU. Version of LSL_ITASK Interface doesn't support multicore");
    return;

  //Check if coreselect is supported by HwControl already
  elsif ( us_CoreSelect > TASK_SELECT_COREMAX ) then
    retcode := -6;
    HWC_LogValue2(this, "@0153 (HwControl::AddHwObject) Invalid parameter us_CoreSelect 0x{0}. Max. us_CoreSelect by HwControl is 0x{1}",us_CoreSelect,TASK_SELECT_COREMAX);
    return;
  end_if;

  //Check if Rt time is smaller than maintimer
  if ( ud_RtTime_us <> 0 ) & ( ud_RtTime_us < _ClockTicks ) then
    retcode := -7;
    HWC_LogError(this, "@0154 (HwControl::AddHwObject) Parameter ud_RtTime_us is smaller than CPU maintimer !");
    return;

  //Check if Rt time is not a multiple of maintimer
  elsif ( ud_RtTime_us <> 0 ) & (ud_RtTime_us MOD _ClockTicks) <> 0 then
    retcode := -8;
    HWC_LogError(this, "@0155 (HwControl::AddHwObject) Parameter ud_RtTime_us not a multiple of CPU maintimer!");
    return;
  end_if;

  //Check if Cy time is smaller than maintimer
  if ( ud_CyTime_us <> 0 ) & ud_CyTime_us < _ClockTicks then
    retcode := -9;
    HWC_LogError(this, "@0156 (HwControl::AddHwObject) Parameter ud_CyTime_us is smaller than CPU maintimer !");
    return;

  //Check if CY time is not a multiple of maintimer
  elsif ( ud_CyTime_us <> 0 ) & (ud_CyTime_us MOD _ClockTicks) <> 0 then
    retcode := -10;
    HWC_LogError(this, "@0157 (HwControl::AddHwObject) Parameter ud_CyTime_us not a multiple of CPU maintimer!");
    return;
  end_if;

  if pHwControlLogins = NIL then
    pHwControlLogins$pVoid := To_StdLib.Malloc(size:=sizeof(t_HwObjectListElement));
    pHelp := pHwControlLogins;
  else
    pHelp := pHwControlLogins;
    while (pHelp^.pThis <> pThis) & (pHelp^.pNext <> NIL) do
      pHelp := pHelp^.pNext;
    end_while;
    if (pHelp^.pThis <> pThis) then
      pHelp^.pNext$pVoid := To_StdLib.Malloc(size:=sizeof(t_HwObjectListElement));
      pHelp := pHelp^.pNext;
//  else
//    already in list and pHelp points to it to update the settings
    end_if;
  end_if;

  if pHelp <> NIL then
    pHelp^.pThis          := pThis;
    pHelp^.pRtPostScan    := NIL;
    pHelp^.bdSettings     := Settings;
    pHelp^.usEscSequence  := EscapeSequence;
    pHelp^.us_CoreSelect  := us_CoreSelect;
    pHelp^.ud_RtTime_us   := ud_RtTime_us;
    pHelp^.ud_CyTime_us   := ud_CyTime_us;
    pHelp^.pNext          := NIL;
    retcode               := 0;
  else
    retcode               := -1;
    HWC_LogError(this,"@015F (HwControl::AddHwObject) Failed to allocate memory for hw object.");
  end_if;

END_FUNCTION

FUNCTION HwControl::PostScanWork
  VAR_INPUT
    us_CoreSelect 	: USINT;
  END_VAR
  VAR
    pHelp : ^t_HwObjectListElement;
#ifdef HWCONTROL_TIME_MEASUREMENT
  udTimeMeasure1 : UDINT;
  udTimeMeasure2 : UDINT;
#endif
  END_VAR

#ifdef HWCONTROL_TIME_MEASUREMENT
  OS_MakeTraceEntry(pSystrace, HWCONTROL_SYSTRACE_TYPE, HWCONTROL_SYSTRACE_RTPOSTSCAN_START,us_CoreSelect);
#endif

  if State = _ClassOk then

    // objects, which are controlled by HwControl (call before the other hardware classes because the safety manager may start moving the data to another system)
    //**********************************************************************************************************************************************************
#ifdef HWCONTROL_TIME_MEASUREMENT
    OS_MakeTraceEntry(pSystrace, HWCONTROL_SYSTRACE_TYPE, HWCONTROL_SYSTRACE_RTPOSTSCAN_START_HW_OBJECTS,us_CoreSelect);
    udTimeMeasure1 := OS_READMICROSEC();
#endif

    UpdateRtPostscanLoginObjects(usCoreSelect:= us_CoreSelect);

#ifdef HWCONTROL_TIME_MEASUREMENT
    udTimeMeasure2 := OS_READMICROSEC();
    aHwControl_Times[us_CoreSelect].sRtPostscan_HwObjects.ActTime := udTimeMeasure2 - udTimeMeasure1;
#endif

    //Call RT Postscan of Varanmanagers
    //**********************************************************************************************************************************************************
#ifdef HWCONTROL_TIME_MEASUREMENT
    OS_MakeTraceEntry(pSystrace, HWCONTROL_SYSTRACE_TYPE, HWCONTROL_SYSTRACE_RTPOSTSCAN_START_VARAN_MANAGERS,us_CoreSelect);
    udTimeMeasure1 := OS_READMICROSEC();
#endif

    UpdateRtPostScanVaranManager(us_CoreSelect);

#ifdef HWCONTROL_TIME_MEASUREMENT
    udTimeMeasure2 := OS_READMICROSEC();
    aHwControl_Times[us_CoreSelect].sRtPostscan_Varan.ActTime := udTimeMeasure2 - udTimeMeasure1;
#endif

  //-------------------------------------Profiler Start----------------------------------------------
  #ifdef	DiasMasterC_Profiler
    HWC_Time_RTPostscan.start := OS_ReadMicroSec();
    if ( ( HWC_Time_RTPostscan.start - HWC_Time_RTPostscan.init ) > DM_ProfilerDelay ) then
      HWC_Time_RTPostscan.initfl := 0;
    else
      HWC_Time_RTPostscan.initfl := 1;
    end_if;
  #endif
  //-------------------------------------Profiler End------------------------------------------------

    if us_CoreSelect = TASK_SELECT_CORE0 then

      if s_DiasMaster.p_Functions <> NIL then
        if s_DiasMaster.p_Functions^.p_RtPostScanFunction <> NIL then
          CallPtr	( p_function := s_DiasMaster.p_Functions^.p_RtPostScanFunction
                  , p_this     := s_DiasMaster.p_Functions^.p_This
                  );
        end_if;
      end_if;

    //Special objects (objects added via the method AddSpecialHW) only run on core 0
      // special classes, which are controlled by HwControl
      if pSpecialObjects then
        pHelp := pSpecialObjects;
        while pHelp <> NIL do
          pHelp^.pRtPostScan$RtWork((pHelp^.pThis)$UDINT);
          pHelp := pHelp^.pNext;
        end_while;
      end_if;
    end_if;

  //-------------------------------------Profiler Stop----------------------------------------------
  #ifdef DiasMasterC_Profiler
    if ( HWC_Time_RTPostscan.initfl = 0 ) then

      HWC_Time_RTPostscan.stop := OS_ReadMicroSec();
      HWC_Time_RTPostscan.diff := HWC_Time_RTPostscan.stop - HWC_Time_RTPostscan.start - DM_CPUconstant;
      HWC_Time_RTPostscan.sum += HWC_Time_RTPostscan.diff;
      HWC_Time_RTPostscan.run += 1;

      if ( HWC_Time_RTPostscan.diff < HWC_Time_RTPostscan._min ) then
        HWC_Time_RTPostscan._min := HWC_Time_RTPostscan.diff;
      end_if;

      if ( HWC_Time_RTPostscan.diff > HWC_Time_RTPostscan._max ) then
        HWC_Time_RTPostscan._max := HWC_Time_RTPostscan.diff;
      end_if;

      HWC_Time_RTPostscan.avg := HWC_Time_RTPostscan.sum * 100 / HWC_Time_RTPostscan.run;

    end_if;
  #endif
  //-------------------------------------Profiler End------------------------------------------------

  end_if;

#ifdef HWCONTROL_TIME_MEASUREMENT
  OS_MakeTraceEntry(pSystrace, HWCONTROL_SYSTRACE_TYPE, HWCONTROL_SYSTRACE_RTPOSTSCAN_FINISH,us_CoreSelect);
  CalcTimeMeasurementPostScan(pHwControlTimes:=#aHwControl_Times[us_CoreSelect]);
#endif

END_FUNCTION

#pragma warning(disable: 73)
FUNCTION VIRTUAL GLOBAL HwControl::AddSafetyManager
  VAR_INPUT
    pThis 	  : pVirtualBase;
  END_VAR
  VAR_OUTPUT
    pFirstVM 	: pVirtualBase;
  END_VAR
#pragma warning(default: 73)

// NO LONGER USED SINCE HWCONTROL HAS IT'S OWN CYCLIC TASK
  pFirstVM := NIL;

END_FUNCTION

FUNCTION VIRTUAL GLOBAL HwControl::SafetyState::Read
  VAR_OUTPUT
    output (EAX) 	: DINT;
  END_VAR

  SafetyState := SafetyManager.ClassState.Read();
  output      := SafetyState;

END_FUNCTION

FUNCTION VIRTUAL GLOBAL HwControl::DisableSafetyManager

// NO LONGER USED SINCE HWCONTROL HAS IT'S OWN CYCLIC TASK

END_FUNCTION

FUNCTION VIRTUAL GLOBAL HwControl::Control::NewInst
  VAR_INPUT
    pPara 	            : ^CmdStruct;
    pResult 	          : ^Results;
  END_VAR
  VAR_OUTPUT
    ret_code 	          : IprStates;
  END_VAR
  VAR
    StartTime                 : UDINT;
    pOneManager               : ^t_OneVaranManager;
    i                         : DINT;
    j                         : DINT;
    TempRetCode               : IprStates;
    MyPara                    : CmdStruct;
    MyResult                  : results;
    pHelp                     : ^t_HwObjectListElement;
    pHelpFirst                : ^t_HwObjectListCallFirst;
    TempSettings              : t_HwObjListSettings;
    us_ModuleType             : HSINT;
    us_CoreSelect             : USINT;
    pStr_HWTRequested         : ^CHAR;
    pStr_HWTreeEntry          : ^CHAR;
    usVaranManagerNrTreeEntry : USINT;
    ud_RtTime_us              : UDINT;
    ud_CyTime_Us              : UDINT;
    sd_retval                 : DINT;
    s_objinfo 		            : LSLOBJ_INFO;
  END_VAR

  us_ModuleType     := 0;
  pStr_HWTRequested := NIL;
  pStr_HWTreeEntry  := NIL;

  ret_code := READY;

  case pPara^.uiCmd of
//**********************************************************************************************************************************************************
    CMD_POST_INIT_CALL:
